(* IEC 61131-3 sources: iecf/harness/cases (part 2) *)

(* ---- enobody.st ---- *)
(* ENO set in a POU's own body (Ed.3 6.6.1.5 rules 2, 3 and 7;
   docs/dependencies.md): ENO is there in every FUNCTION and
   FUNCTION_BLOCK without a declaration, TRUE as each run starts, and the
   caller's ENO is FALSE when the body set it FALSE or a flag was raised
   while it ran. `lim` clears ENO above 100, `half` below 0; `acc` sets
   ENO TRUE at its end, which cannot hide the overflow of its fifth run
   (tick 4): iecf's ENO is FALSE there, the reference compiler's TRUE, as
   it has no flag; iecf's trace is enobody.iecf.trace. The input v is
   5, 200, -4, 30000, 30000. r_bits: bit 0 lim's ENO, 1 half's, 2 acc's. *)
FUNCTION_BLOCK lim
VAR_INPUT x : INT; END_VAR
VAR_OUTPUT y : INT; END_VAR
y := x;
IF x > 100 THEN ENO := FALSE; END_IF;
END_FUNCTION_BLOCK

FUNCTION half : INT
VAR_INPUT x : INT; END_VAR
half := x / 2;
ENO := x >= 0;
END_FUNCTION

FUNCTION_BLOCK acc
VAR_INPUT x : INT; END_VAR
VAR_OUTPUT total : INT; END_VAR
total := total + x;
ENO := TRUE;
END_FUNCTION_BLOCK

PROGRAM main
VAR
  v AT %IW0 : INT;
  r_bits AT %MB0 : BYTE;
  r_half AT %MB1 : SINT;
  r_y AT %MW2 : INT;
  r_total AT %MW4 : INT;
END_VAR
VAR
  l : lim;
  a : acc;
  ok1, ok2, ok3 : BOOL;
  h : INT;
END_VAR
l(x := v, y => r_y, ENO => ok1);
h := half(x := v, ENO => ok2);
r_half := INT_TO_SINT(h / 1000);
a(x := v, total => r_total, ENO => ok3);
r_bits := 0;
IF ok1 THEN r_bits := r_bits OR 16#01; END_IF;
IF ok2 THEN r_bits := r_bits OR 16#02; END_IF;
IF ok3 THEN r_bits := r_bits OR 16#04; END_IF;
END_PROGRAM

CONFIGURATION plant
  RESOURCE r ON PLC
    TASK fast(INTERVAL := T#10ms, PRIORITY := 0);
    PROGRAM p WITH fast : main;
  END_RESOURCE
END_CONFIGURATION

(* ---- enointo.st ---- *)
(* A block's ENO, and outputs, taken into an element, a field and a bit,
   each found - its index checked - before the block runs. Worked by
   hand:
   t(EN := TRUE, ..., ENO => a[i]), i 2: ENO TRUE, a[2] TRUE (%QX0.0).
   t(EN := FALSE, ..., NOT ENO => w.3): ENO FALSE, its NOT TRUE: w 8,
   w.%B0 08 (%QB1).
   t(EN := TRUE, ..., ENO => s.ok): s.ok TRUE (%QX0.1).
   o(q => ws[i].3, qb => ws[i].%B1), q TRUE and qb 7: ws[2] 16#0708,
   its bytes 08 (%QB2) and 07 (%QB3).
   F(q => ws[1].2), q TRUE: ws[1] 4 (%QB4).
   Last, i 3: o(q => ws[i].0) faults (INDEX) before o runs, so n, o's
   count of its runs, stays 1 (%QB5).
   reference-skip: partial access, NOT ENO =>: refused (iec2c crashes
   on the latter). *)
TYPE
  STV : STRUCT ok : BOOL; END_STRUCT;
END_TYPE
FUNCTION_BLOCK OT
  VAR_OUTPUT q : BOOL; qb : BYTE; n : INT; END_VAR
  q := TRUE;
  qb := 7;
  n := n + 1;
END_FUNCTION_BLOCK
FUNCTION F : INT
  VAR_OUTPUT q : BOOL; END_VAR
  q := TRUE;
  F := 1;
END_FUNCTION
PROGRAM main
  VAR
    t : TON;
    o : OT;
    a : ARRAY [1..2] OF BOOL;
    ws : ARRAY [1..2] OF WORD;
    s : STV;
    w : WORD;
    i : INT := 2;
    v : INT;
  END_VAR
  VAR
    q00 AT %QX0.0 : BOOL;
    q01 AT %QX0.1 : BOOL;
    q1 AT %QB1 : BYTE;
    q2 AT %QB2 : BYTE;
    q3 AT %QB3 : BYTE;
    q4 AT %QB4 : BYTE;
    q5 AT %QB5 : SINT;
  END_VAR
  t(EN := TRUE, IN := FALSE, PT := T#1s, ENO => a[i]);
  q00 := a[2];
  t(EN := FALSE, IN := FALSE, PT := T#1s, NOT ENO => w.3);
  q1 := w.%B0;
  t(EN := TRUE, IN := FALSE, PT := T#1s, ENO => s.ok);
  q01 := s.ok;
  o(q => ws[i].3, qb => ws[i].%B1);
  q2 := ws[2].%B0;
  q3 := ws[2].%B1;
  v := F(q => ws[1].2);
  q4 := ws[1].%B0;
  q5 := INT_TO_SINT(o.n);
  i := 3;
  o(q => ws[i].0);
END_PROGRAM

CONFIGURATION c
  RESOURCE r ON x
    TASK t(INTERVAL := T#10ms, PRIORITY := 1);
    PROGRAM p WITH t : main;
  END_RESOURCE
END_CONFIGURATION

(* ---- enums.st ---- *)
(* Enumerations and types with named values (Ed.3 6.4.4.2, 6.4.4.3).
   col has named values: red 1, green 5, blue one more, 6; its initial
   value green. A col is used as the INT it is: other values assigned,
   arithmetic, comparison. mode is an enumeration, its initial value run.
   An enumeration is a FUNCTION's input, output and result and a block's
   in-out; a result or an input not given starts as the type's initial
   value. Worked by hand, k %IB0 1, 2, 3:
   %QB0: c as the tick starts: 5 (green), then what the tick before left,
   3, 4. %QB1: x := c + blue when c = green: 11, and kept.
   c := k, then CASE c OF red: 10; green - 3 (2), blue: 20; ELSE 30:
   %QB2 10, 20, 30.
   b(c := c, m := m, d := red + 1): c + 2, %QB3 3, 4, 5; m := NEXT(m):
   run gives stop; stop matches no label, so NEXT keeps its initial value,
   run; then stop again: %QB4 2, 1, 2 (stop 2, run 1).
   lv#hi OR lo, a WORD: 16#30, %QB5.
   n, an INT, given to the in-out c: 10 + blue each tick: %QB6 16, 22, 28.
   m3 := DEF(o => m4), both idle before: DEF's result is not set and its
   input m not given, so both are run: %QB7 1.
   %QB8 blue, 6. %QB9 a[2], an array's element of col: green, 5.
   mi : (low, mid, top) := mid, declared in place: mid gives 7 and
   becomes top, top gives 8: %QB10 7, 8, 8.
   gear names no base type, so it is an INT (as CODESYS and TwinCAT
   have it) and is added to one as it is: g is slow, 2; x2, an INT from
   3, x2 := x2 + g each tick: %QB11 5, 7, 9.
   reference-skip: named values are Ed.3's; the reference compiler
   (Ed.2) has none. *)
TYPE
  col : INT (red := 1, green := 5, blue) := green;
  lv : WORD (lo := 16#10, hi := 16#20);
  mode : (idle, run, stop) := run;
  gear : (slow := 2, fast := 4);
END_TYPE

FUNCTION NEXT : mode
  VAR_INPUT m : mode; END_VAR
  CASE m OF
    idle: NEXT := run;
    run: NEXT := stop;
  END_CASE;
END_FUNCTION

FUNCTION DEF : mode
  VAR_INPUT m : mode; END_VAR
  VAR_OUTPUT o : mode; END_VAR
  o := m;
END_FUNCTION

FUNCTION_BLOCK BUMP
  VAR_IN_OUT c : col; m : mode; END_VAR
  VAR_INPUT d : col; END_VAR
  c := c + d;
  m := NEXT(m);
END_FUNCTION_BLOCK

PROGRAM main
  VAR
    c : col;
    x : INT;
    w : WORD;
    m, m2 : mode;
    m3, m4 : mode := idle;
    b : BUMP;
    n : INT := 10;
    a : ARRAY [1..2] OF col;
    mi : (low, mid, top) := mid;
    g : gear;
    x2 : INT := 3;
  END_VAR
  VAR k AT %IB0 : SINT; END_VAR
  VAR
    q0 AT %QB0 : SINT;
    q1 AT %QB1 : SINT;
    q2 AT %QB2 : SINT;
    q3 AT %QB3 : SINT;
    q4 AT %QB4 : SINT;
    q5 AT %QB5 : BYTE;
    q6 AT %QB6 : SINT;
    q7 AT %QB7 : SINT;
    q8 AT %QB8 : SINT;
    q9 AT %QB9 : SINT;
    q10 AT %QB10 : SINT;
    q11 AT %QB11 : SINT;
  END_VAR
  q0 := INT_TO_SINT(c);
  IF c = col#green THEN
    x := c + blue;
  END_IF;
  q1 := INT_TO_SINT(x);
  c := k;
  CASE c OF
    red: q2 := 10;
    green - 3, blue: q2 := 20;
  ELSE
    q2 := 30;
  END_CASE;
  b(c := c, m := m, d := red + 1);
  q3 := INT_TO_SINT(c);
  IF m = stop THEN
    q4 := 2;
  ELSIF m = mode#run THEN
    q4 := 1;
  ELSE
    q4 := 0;
  END_IF;
  w := lv#hi OR lo;
  q5 := WORD_TO_BYTE(w);
  b(c := n, m := m2, d := blue);
  q6 := INT_TO_SINT(n);
  m3 := DEF(o => m4);
  IF m3 = run AND m4 = run THEN
    q7 := 1;
  END_IF;
  q8 := INT_TO_SINT(blue);
  q9 := INT_TO_SINT(a[2]);
  IF mi = mid THEN
    q10 := 7;
    mi := top;
  ELSIF mi = top THEN
    q10 := 8;
  END_IF;
  x2 := x2 + g;
  q11 := INT_TO_SINT(x2);
END_PROGRAM

CONFIGURATION c
  RESOURCE r ON PLC
    TASK t(INTERVAL := T#10ms, PRIORITY := 1);
    PROGRAM p WITH t : main;
  END_RESOURCE
END_CONFIGURATION

(* ---- fbargs.st ---- *)
(* A function block's in-out given, and its output taken into, any
   variable of the type (Ed.3 6.6.3.4): an element by a constant and by
   a computed index, a field, a variable through a reference, an
   element at an address. And an enumeration declared in place with
   named values (Ed.3 6.4.4.3), used as its base type.
   ADD1 adds 1 to its in-out v; twice := 2 * v; neg := v < 0.
   Worked by hand, k %IB0 1, 2, 3; arr and out start [0, 0, 0]:
   b(v := arr[2], twice => out[1]); i := k; b(v := arr[i], twice =>
   out[i]); and, last in the scan, b(v := arr[k + 1]):
     tick 0: arr[2] 1, out[1] 2; i 1: arr[1] 1, out[1] 2; arr [1, 1,
     0], out [2, 0, 0]; then arr[2] 2.
     tick 1: arr[2] 3, out[1] 6; i 2: arr[2] 4, out[2] 8; arr [1, 4,
     0], out [6, 8, 0]; then arr[3] 1.
     tick 2: arr[2] 5, out[1] 10; i 3: arr[3] 2, out[3] 4; arr [1, 5,
     2], out [10, 8, 4]; then arr[4], outside 1..3: a fault (index),
     before the block runs.
     %QB0..2 arr, %QB3..5 out.
   b(v := p.y, twice => po.x): p.y 1, 2, 3 (%QB6); po.x 2, 4, 6 (%QB7).
   b(v := r^, twice => ro^), r to tgt, ro to d2: tgt + 1, d2 twice it.
   b(v := tgt, twice => d), d a DINT, the output widened: tgt + 1
   again: tgt 2, 4, 6 (%QB8); d2 2, 6, 10 (%QB9); d 4, 8, 12 (%QB10).
   b(v := p.x, NOT neg => nb): nb TRUE (%QX11.0).
   b(v := lm[2], twice => lm[1]), lm at %MW0: lm[2] 1, 2, 3 and lm[1]
   2, 4, 6 in %MW2 and %MW0.
   x : INT (lo := 1, hi := 5) := hi, in place: x + lo 6, then x := x + 1:
   6, 7, 8 (%QB12). y : (p3 := 3, q4): 3, then y := q4: 3, 4, 4 (%QB13).
   SPARE is a block with an instance that is never called: the C still
   builds with every warning an error, as the harness builds it.
   reference-skip: named values are Ed.3's; the reference compiler
   (Ed.2) has none. *)
TYPE PT : STRUCT x, y : INT; END_STRUCT; END_TYPE
FUNCTION_BLOCK ADD1
  VAR_IN_OUT v : INT; END_VAR
  VAR_OUTPUT twice : INT; neg : BOOL; END_VAR
  v := v + 1;
  twice := 2 * v;
  neg := v < 0;
END_FUNCTION_BLOCK
FUNCTION_BLOCK SPARE
  VAR_INPUT a : INT; END_VAR
  VAR_OUTPUT o : INT; END_VAR
  o := a;
END_FUNCTION_BLOCK
CONFIGURATION c
  RESOURCE r ON PLC
    TASK t(INTERVAL := T#10ms, PRIORITY := 1);
    PROGRAM p WITH t : main;
  END_RESOURCE
END_CONFIGURATION
PROGRAM main
  VAR
    arr, out : ARRAY [1..3] OF INT;
    p, po : PT;
    r, ro : REF_TO INT;
    tgt, d2, i : INT;
    d : DINT;
    nb : BOOL;
    b : ADD1;
    idle : SPARE;
    x : INT (lo := 1, hi := 5) := hi;
    y : (p3 := 3, q4);
  END_VAR
  VAR lm AT %MW0 : ARRAY [1..2] OF INT; END_VAR
  VAR k AT %IB0 : SINT; END_VAR
  VAR
    q0 AT %QB0 : SINT;
    q1 AT %QB1 : SINT;
    q2 AT %QB2 : SINT;
    q3 AT %QB3 : SINT;
    q4b AT %QB4 : SINT;
    q5 AT %QB5 : SINT;
    q6 AT %QB6 : SINT;
    q7 AT %QB7 : SINT;
    q8 AT %QB8 : SINT;
    q9 AT %QB9 : SINT;
    q10 AT %QB10 : SINT;
    q11 AT %QX11.0 : BOOL;
    q12 AT %QB12 : SINT;
    q13 AT %QB13 : SINT;
  END_VAR
  b(v := arr[2], twice => out[1]);
  i := k;
  b(v := arr[i], twice => out[i]);
  b(v := p.y, twice => po.x);
  r := REF(tgt);
  ro := REF(d2);
  b(v := r^, twice => ro^);
  b(v := tgt, twice => d);
  b(v := p.x, NOT neg => nb);
  b(v := lm[2], twice => lm[1]);
  q0 := INT_TO_SINT(arr[1]);
  q1 := INT_TO_SINT(arr[2]);
  q2 := INT_TO_SINT(arr[3]);
  q3 := INT_TO_SINT(out[1]);
  q4b := INT_TO_SINT(out[2]);
  q5 := INT_TO_SINT(out[3]);
  q6 := INT_TO_SINT(p.y);
  q7 := INT_TO_SINT(po.x);
  q8 := INT_TO_SINT(tgt);
  q9 := INT_TO_SINT(d2);
  q10 := DINT_TO_SINT(d);
  q11 := nb;
  q12 := INT_TO_SINT(x + lo);
  x := x + 1;
  q13 := INT_TO_SINT(y);
  y := q4;
  b(v := arr[k + 1]);
END_PROGRAM

(* ---- fbeffects.st ---- *)
(* FUNCTIONs with effects in a block call: in the index of the target an
   output is taken into, and as a STRING input. Each is made once, in
   order; an output's target is found after the block runs, as a
   FUNCTION's is, so a call there runs after the block does
   (docs/dependencies.md). Worked by hand, each tick from j 1:

   f(io := j, s := 'x', q => a[finc(j)]): the block, io j 1: q 1 +
   LEN('x') 1 = 2; then finc makes j 2 and gives 2, the target a[2]:
   2 (Q0 02). f(io := j, s := fso(x := 'bb', y => j)): fso gives
   'bb' and sets j to 7; then the block, io 7: q 7 + 2 = 9 (Q1 09); j 7
   (Q2 07).
   fbeffects.iecf.trace: the reference compiler copies the in-out in
   before the other inputs are computed and back after the call, so
   fso's j is lost (Q 02 04 02); iecf binds the in-out to j itself. *)
FUNCTION finc : INT
  VAR_IN_OUT x : INT; END_VAR
  x := x + 1;
  finc := x;
END_FUNCTION
FUNCTION fso : STRING
  VAR_INPUT x : STRING; END_VAR
  VAR_OUTPUT y : INT; END_VAR
  y := 7;
  fso := x;
END_FUNCTION
FUNCTION_BLOCK fb
  VAR_IN_OUT io : INT; END_VAR
  VAR_INPUT s : STRING; END_VAR
  VAR_OUTPUT q : INT; END_VAR
  q := io + LEN(s);
END_FUNCTION_BLOCK
PROGRAM main
  VAR f : fb; a : ARRAY [1..4] OF INT; j : INT; END_VAR
  VAR q AT %QB0 : USINT; q1 AT %QB1 : USINT; q2 AT %QB2 : USINT; END_VAR
  j := 1;
  f(io := j, s := 'x', q => a[finc(j)]);
  q := INT_TO_USINT(a[2]);
  f(io := j, s := fso(x := 'bb', y => j));
  q1 := INT_TO_USINT(f.q);
  q2 := INT_TO_USINT(j);
END_PROGRAM
CONFIGURATION c RESOURCE r ON PLC TASK t(INTERVAL := T#10ms, PRIORITY := 1); PROGRAM p WITH t : main; END_RESOURCE END_CONFIGURATION

(* ---- fbenable.st ---- *)
(* EN and ENO on a function block call (Ed.3 6.6.1.5; docs/dependencies.md):
   an accumulator adds 10000 at each call it is enabled for, %IX0.0 its EN.
   Each tick r_n is set to -1 before the call: with EN FALSE (tick 1) the
   block is not called, its total stays and is not taken into r_n, and ENO
   is FALSE. Its fourth enabled call (tick 4) overflows inside the block:
   the total wraps, the flag is raised in the block's body, and ENO is
   FALSE. r_bits: bit 0 ENO. The reference compiler takes the output into
   r_n with EN FALSE and has no flag to clear ENO: iecf's trace is
   fbenable.iecf.trace. NOT ENO, which the reference compiler cannot
   compile, is fbskip's. *)
FUNCTION_BLOCK acc
VAR_INPUT x : INT; END_VAR
VAR_OUTPUT total : INT; END_VAR
total := total + x;
END_FUNCTION_BLOCK

PROGRAM main
VAR
  c AT %IX0.0 : BOOL;
  r_n AT %MW0 : INT;
  r_total AT %MW2 : INT;
  r_bits AT %MB4 : BYTE;
END_VAR
VAR
  a : acc;
  ok : BOOL;
END_VAR
r_n := -1;
a(EN := c, x := 10000, total => r_n, ENO => ok);
r_total := a.total;
r_bits := 0;
IF ok THEN r_bits := r_bits OR 16#01; END_IF;
END_PROGRAM

CONFIGURATION plant
  RESOURCE r ON PLC
    TASK fast(INTERVAL := T#10ms, PRIORITY := 0);
    PROGRAM p WITH fast : main;
  END_RESOURCE
END_CONFIGURATION

(* ---- fbencall.st ---- *)
(* A function block's EN given a call (Ed.3 6.6.1.5): of a FUNCTION
   with an in-out, of a method, of a method through an interface. EN is
   computed first, once, and only then the block is called or not, ENO
   telling which. Worked by hand, tick by tick:
   Advance adds 1 to n and gives n > 2: n 1, 2, 3, 4; c1 runs at ticks
   2 and 3, total (%QB0) 0, 0, 1, 2; n (%QB1); ENO e1 (%QX4.0) FALSE,
   FALSE, TRUE, TRUE.
   v.Ready gives its count < 2, then counts: TRUE, TRUE, FALSE, FALSE;
   c2 adds 10: 10, 20, 20, 20 (%QB2); e2 (%QX4.1).
   ig.Open counts and gives whether its count is even: FALSE, TRUE,
   FALSE, TRUE; c3 adds 5: 0, 5, 5, 10 (%QB3); e3 (%QX4.2).
   reference-skip: METHOD and INTERFACE are Ed.3's; the reference
   compiler (Ed.2) has neither. *)
FUNCTION Advance : BOOL
  VAR_IN_OUT cnt : INT; END_VAR
  cnt := cnt + 1;
  Advance := cnt > 2;
END_FUNCTION

FUNCTION_BLOCK Valve
  VAR n : INT; END_VAR
  METHOD PUBLIC Ready : BOOL
    Ready := n < 2;
    n := n + 1;
  END_METHOD
END_FUNCTION_BLOCK

INTERFACE IGate
  METHOD Open : BOOL
  END_METHOD
END_INTERFACE

FUNCTION_BLOCK Gate IMPLEMENTS IGate
  VAR k : INT; END_VAR
  METHOD PUBLIC Open : BOOL
    k := k + 1;
    Open := k MOD 2 = 0;
  END_METHOD
END_FUNCTION_BLOCK

FUNCTION_BLOCK Count
  VAR_INPUT inc : INT; END_VAR
  VAR_OUTPUT total : INT; END_VAR
  total := total + inc;
END_FUNCTION_BLOCK

PROGRAM main
  VAR
    n : INT;
    v : Valve;
    g : Gate;
    ig : IGate;
    c1, c2, c3 : Count;
  END_VAR
  VAR
    q0 AT %QB0 : SINT;
    q1 AT %QB1 : SINT;
    q2 AT %QB2 : SINT;
    q3 AT %QB3 : SINT;
    e1 AT %QX4.0 : BOOL;
    e2 AT %QX4.1 : BOOL;
    e3 AT %QX4.2 : BOOL;
  END_VAR
  ig := g;
  c1(EN := Advance(n), inc := 1, ENO => e1);
  c2(EN := v.Ready(), inc := 10, ENO => e2);
  c3(EN := ig.Open(), inc := 5, ENO => e3);
  q0 := INT_TO_SINT(c1.total);
  q1 := INT_TO_SINT(n);
  q2 := INT_TO_SINT(c2.total);
  q3 := INT_TO_SINT(c3.total);
END_PROGRAM

CONFIGURATION c
  RESOURCE r ON x
    TASK t(INTERVAL := T#10ms, PRIORITY := 1);
    PROGRAM p WITH t : main;
  END_RESOURCE
END_CONFIGURATION

(* ---- fbinitarrays.st ---- *)
(* CODESYS's and TwinCAT's arrays of instances set up by their FB_init
   (fb-init), as TcOpen's `ARRAY[0..2] OF DiagnosticsMessenger(THIS^)`,
   and in-outs of a type with an FB_init, bound, not set up.
   Worked by hand: h's items, its first VAR, are set up first, each
   element's FB_init in index order given THIS^, h: each takes h.Next(),
   1 2 3; then grid, row by row, (1,-1) (1,0) (2,-1) (2,0): 4 5 6 7;
   then plain, with no arguments, each element's FB_init counting itself
   once, bInitRetains TRUE at the cold start; then d, a structure whose
   member cells is such an array, then nest, an array of arrays.
   %QW0 items[0..2] 1 2 3 as 123, %QW2 grid as 4567, %QW4 h.seq 7,
   %QW6 plain's counts summed, 3, %QW8 those cold, 3, %QW10 d.cells'
   counts summed, 2, and nest's, 4, times 10: 42; %QW12 h.u reading items[2] through its in-out, 3,
   %QW14 its method reading grid[2, 0] through one, 7.
   reference-skip: not IEC 61131-3. *)
INTERFACE ISeq
  METHOD Next : INT
  END_METHOD
END_INTERFACE

FUNCTION_BLOCK Item
  VAR_OUTPUT mine : INT; END_VAR
  METHOD FB_init : BOOL
    VAR_INPUT bInitRetains : BOOL; bInCopyCode : BOOL; s : ISeq; END_VAR
    mine := s.Next();
  END_METHOD
END_FUNCTION_BLOCK

FUNCTION_BLOCK Counted
  VAR_OUTPUT times : INT; cold : INT; END_VAR
  METHOD FB_init : BOOL
    VAR_INPUT bInitRetains : BOOL; bInCopyCode : BOOL; END_VAR
    times := times + 1;
    IF bInitRetains THEN cold := cold + 1; END_IF
  END_METHOD
END_FUNCTION_BLOCK

TYPE Cells : STRUCT
  tag : INT := 1;
  cells : ARRAY[0..1] OF Counted;
END_STRUCT
END_TYPE

FUNCTION_BLOCK User
  VAR_IN_OUT io : Item; END_VAR
  VAR_OUTPUT o : INT; END_VAR
  METHOD Read : INT
    VAR_IN_OUT other : Item; END_VAR
    Read := other.mine;
  END_METHOD
  o := io.mine;
END_FUNCTION_BLOCK

FUNCTION_BLOCK Holder IMPLEMENTS ISeq
  VAR
    seq : INT;
    items : ARRAY[0..2] OF Item(THIS^);
    grid : ARRAY[1..2, -1..0] OF Item(THIS^);
    plain : ARRAY[0..2] OF Counted;
    d : Cells;
    nest : ARRAY[0..1] OF ARRAY[0..1] OF Counted;
    u : User;
  END_VAR
  VAR_OUTPUT o1 : INT; o2 : INT; o3 : INT; o4 : INT; o5 : INT; o6 : INT; o7 : INT; o8 : INT; END_VAR
  VAR_TEMP k : INT; END_VAR
  METHOD PUBLIC Next : INT
    seq := seq + 1;
    Next := seq;
  END_METHOD
  o1 := items[0].mine * 100 + items[1].mine * 10 + items[2].mine;
  o2 := grid[1, -1].mine * 1000 + grid[1, 0].mine * 100 + grid[2, -1].mine * 10 + grid[2, 0].mine;
  o3 := seq;
  o4 := 0; o5 := 0;
  FOR k := 0 TO 2 DO
    o4 := o4 + plain[k].times;
    o5 := o5 + plain[k].cold;
  END_FOR
  o6 := d.cells[0].times + d.cells[1].times;
  FOR k := 0 TO 1 DO
    o6 := o6 + 10 * (nest[k][0].times + nest[k][1].times);
  END_FOR
  u(io := items[2]);
  o7 := u.o;
  o8 := u.Read(other := grid[2, 0]);
END_FUNCTION_BLOCK

PROGRAM main
  VAR h : Holder; END_VAR
  VAR q0 AT %QW0 : INT; q1 AT %QW2 : INT; q2 AT %QW4 : INT; q3 AT %QW6 : INT; q4 AT %QW8 : INT;
      q5 AT %QW10 : INT; q6 AT %QW12 : INT; q7 AT %QW14 : INT; END_VAR
  h();
  q0 := h.o1; q1 := h.o2; q2 := h.o3; q3 := h.o4; q4 := h.o5; q5 := h.o6;
  q6 := h.o7; q7 := h.o8;
END_PROGRAM

CONFIGURATION cf
  RESOURCE r ON x
    TASK tk(INTERVAL := T#10ms, PRIORITY := 1);
    PROGRAM p WITH tk : main;
  END_RESOURCE
END_CONFIGURATION

(* ---- fbinorder.st ---- *)
(* A function block called with its arguments in order (Ed.3 6.6.3.4.1,
   the non-formal call): every input, output and in-out where it is
   declared, a base's first, none left off ("exactly the same number of
   parameters, in exactly the same order", 6.6.1.4.2). Worked by hand:

   tick 0. adder declares a, b, o, n, o2: f(1, 2, r, x, r2) gives a 1,
   b 2, o into r, the in-out n is x, o2 into r2: r 3 (Q0), r2 -1 (Q2 ff
   ff), x 1 (Q4). f(10, 20, r, x, r2): f.o 30 (Q6 1e 00), x 2. g, a
   wider, takes adder's a, b, o, n, o2, then its own c, p, s, o3: g(1,
   2, r, x, r2, 3, pt, 'abc', r3) gives o 3, x 3, o3 3 + 3 + 100 + 3 =
   109 (Q8 6d 00). g.twice(7, h): 14, h 3: 17 (Q10 11 00). TON's IN,
   PT, Q, ET: t(TRUE, T#20ms, done, el): not done (Q12 0); CTU's CU, R,
   PV, Q, CV: ctr(done, FALSE, 5, cq, cv): 0 (Q14).
   tick 1: x was 3: 4 after the first call (Q4 04 00); the rest as
   before.
   tick 2: x 7; t is done after 20 ms (Q12 01 00), and ctr counts its
   rising edge: 1 (Q14).
   tick 3: x 10; done stays, the count stays 1.
   reference-skip: methods, EXTENDS: refused. *)
TYPE PtT : STRUCT x : INT; y : INT; END_STRUCT; END_TYPE
FUNCTION_BLOCK adder
  VAR_INPUT a : INT; b : INT := 5; END_VAR
  VAR_OUTPUT o : INT; END_VAR
  VAR_IN_OUT n : INT; END_VAR
  VAR_OUTPUT o2 : INT; END_VAR
  o := a + b;
  n := n + 1;
  o2 := a - b;
END_FUNCTION_BLOCK
FUNCTION_BLOCK wider EXTENDS adder
  VAR_INPUT c : INT; p : PtT; s : STRING[4]; END_VAR
  VAR_OUTPUT o3 : INT; END_VAR
  METHOD PUBLIC twice : INT
    VAR_INPUT v : INT; END_VAR
    VAR_OUTPUT half : INT; END_VAR
    twice := v * 2;
    half := v / 2;
  END_METHOD
  SUPER();
  o3 := o + c + p.x + LEN(s);
END_FUNCTION_BLOCK
PROGRAM main
  VAR f : adder; g : wider; t : TON; ctr : CTU; x : INT; r, r2, r3, m, h : INT; pt : PtT := (x := 100); el : TIME; done, cq : BOOL; cv : INT; END_VAR
  VAR q AT %QW0 : ARRAY [0..7] OF INT; END_VAR
  f(1, 2, r, x, r2);
  q[0] := r; q[1] := r2; q[2] := x;
  f(10, 20, r, x, r2);
  q[3] := f.o;
  g(1, 2, r, x, r2, 3, pt, 'abc', r3);
  q[4] := r3;
  m := g.twice(7, h);
  q[5] := m + h;
  t(TRUE, T#20ms, done, el);
  q[6] := BOOL_TO_INT(done);
  ctr(done, FALSE, 5, cq, cv);
  q[7] := ctr.CV;
END_PROGRAM
CONFIGURATION c RESOURCE r ON PLC TASK t(INTERVAL := T#10ms, PRIORITY := 1); PROGRAM p WITH t : main; END_RESOURCE END_CONFIGURATION

(* ---- fbparts.st ---- *)
(* A part of a block's elementary input or output read from outside
   (Ed.3 Table 17): `f.q.%X4`, `f.q.%B1`, of an element of an array of
   instances, in a condition. Worked by hand: f.iw 16#0123, so f.q is
   ROL(16#0123, 4), 16#1230: its byte 1 is 16#12 (Q0); its bit 4 is 1,
   iw's bit 1 is 1, fa[2].q is 16#0040 and its bit 6 is 1, f.q's bit 5
   is 1: the four bits 2#1111 (Q1 0f).
   reference-skip: partial access, as `partaccess`. *)
FUNCTION_BLOCK fb
  VAR_INPUT iw : WORD; END_VAR
  VAR_OUTPUT q : WORD; END_VAR
  q := ROL(iw, 4);
END_FUNCTION_BLOCK
PROGRAM main
  VAR f : fb; fa : ARRAY [1..2] OF fb; i : INT := 2; b1, b2, b3, b4 : BOOL; y : BYTE; END_VAR
  VAR q AT %QB0 : BYTE; q1 AT %QB1 : BYTE; END_VAR
  f(iw := 16#0123);
  fa[2](iw := 16#0004);
  b1 := f.q.%X4;
  y := f.q.%B1;
  b2 := f.iw.%X1;
  b3 := fa[i].q.%X6;
  IF f.q.%X5 THEN b4 := TRUE; END_IF;
  q := y;
  q1 := BOOL_TO_BYTE(b1) OR SHL(BOOL_TO_BYTE(b2), 1) OR SHL(BOOL_TO_BYTE(b3), 2) OR SHL(BOOL_TO_BYTE(b4), 3);
END_PROGRAM
CONFIGURATION c RESOURCE r ON PLC TASK t(INTERVAL := T#10ms, PRIORITY := 1); PROGRAM p WITH t : main; END_RESOURCE END_CONFIGURATION

(* ---- fbretain.st ---- *)
(* RETAIN inside a FUNCTION_BLOCK (Ed.3 6.5.6): at a warm restart the
   block's own RETAIN variable keeps its value, its NON_RETAIN one is set
   anew, and one that is neither keeps its value only in an instance
   declared RETAIN. A block in a block follows its own type and the
   section it is declared in, not the outer instance. An instance of a
   block that keeps anything is kept whole (docs/c-output.md §7).
   Each counter counts from 10, 20, 30; at tick 3 a warm restart.
   The reference compiler has no warm restart of its own; its host starts everything
   anew. iecf's trace is fbretain.iecf.trace. *)
FUNCTION_BLOCK cnt
VAR_OUTPUT
  ko : INT;
  po : INT;
  no : INT;
END_VAR
VAR RETAIN
  k : INT := 10;
END_VAR
VAR
  p : INT := 20;
END_VAR
VAR NON_RETAIN
  n : INT := 30;
END_VAR
k := k + 1;
p := p + 1;
n := n + 1;
ko := k;
po := p;
no := n;
END_FUNCTION_BLOCK

FUNCTION_BLOCK wrap
VAR_OUTPUT
  ck, cp, cn, dk, dp, dn : INT;
END_VAR
VAR
  c : cnt;
END_VAR
VAR RETAIN
  cr : cnt;
END_VAR
c();
cr();
ck := c.ko;
cp := c.po;
cn := c.no;
dk := cr.ko;
dp := cr.po;
dn := cr.no;
END_FUNCTION_BLOCK

PROGRAM main
VAR
  a_k AT %MW0 : INT;
  a_p AT %MW2 : INT;
  a_n AT %MW4 : INT;
  b_k AT %MW6 : INT;
  b_p AT %MW8 : INT;
  b_n AT %MW10 : INT;
  c_k AT %MW12 : INT;
  c_p AT %MW14 : INT;
  c_n AT %MW16 : INT;
  d_k AT %MW18 : INT;
  d_p AT %MW20 : INT;
  d_n AT %MW22 : INT;
END_VAR
VAR
  a : cnt;
  w : wrap;
END_VAR
VAR RETAIN
  b : cnt;
END_VAR
a();
b();
w();
a_k := a.ko;
a_p := a.po;
a_n := a.no;
b_k := b.ko;
b_p := b.po;
b_n := b.no;
c_k := w.ck;
c_p := w.cp;
c_n := w.cn;
d_k := w.dk;
d_p := w.dp;
d_n := w.dn;
END_PROGRAM

CONFIGURATION plant
  RESOURCE r ON PLC
    TASK fast(INTERVAL := T#10ms, PRIORITY := 0);
    PROGRAM p WITH fast : main;
  END_RESOURCE
END_CONFIGURATION

(* ---- fbskip.st ---- *)
(* A function block call with EN FALSE is not made at all (Ed.3 6.6.1.5,
   Example 2; docs/dependencies.md): its inputs are not evaluated - x
   divides by zero and nothing faults - nor set, the block does not run,
   its output is not taken, and NOT ENO gives TRUE. With EN TRUE at tick 1
   (zero is 1 by then) it runs once. The reference compiler cannot compile
   `NOT ENO =>` (PROPOSAL.md §1b): iecf only. *)
FUNCTION_BLOCK acc
VAR_INPUT x : INT; END_VAR
VAR_OUTPUT total : INT; END_VAR
total := total + x;
END_FUNCTION_BLOCK

PROGRAM main
VAR
  r_n AT %MW0 : INT;
  r_total AT %MW2 : INT;
  r_off AT %MX4.0 : BOOL;
END_VAR
VAR
  a : acc;
  run : BOOL;
  zero : INT;
END_VAR
r_n := -1;
a(EN := run, x := 100 / zero, total => r_n, NOT ENO => r_off);
r_total := a.total;
run := TRUE;
zero := 1;
END_PROGRAM

CONFIGURATION plant
  RESOURCE r ON PLC
    TASK fast(INTERVAL := T#10ms, PRIORITY := 0);
    PROGRAM p WITH fast : main;
  END_RESOURCE
END_CONFIGURATION

(* ---- flexarrays.st ---- *)
(* Variable-length arrays (Ed.3 6.5.3) and named constants in bounds
   (Ed.3 6.6.1.2.4). SUM is Ed.3's Example 2: it adds an ARRAY[*] whatever
   its bounds. FILL writes a 2-dimensional one, M[i, j] := 10 * i + j.
   TWICE passes its ARRAY[*] on to SUM. A CLASS's method takes one too.
   W, a VAR_GLOBAL CONSTANT, bounds a TYPE; N, the program's own
   CONSTANT, bounds an array and a STRING; a subrange is 0..N.
   Worked by hand, k %IB0:
   a: 1..5 (N), [1, 2, 3, 4, 5]: SUM 15, %QB0 15. b: -2..2, [10, 20, 30,
   40, 50]: SUM 150, %QB1 150. TWICE(a) 2 * 15 = 30, %QB2 30.
   m: 1..2, -1..1 filled: m[1, -1] 9, m[2, 1] 21: %QB3 9, %QB4 21.
   LOWER_BOUND(b, 1) -2, %QB5 16#fe; UPPER_BOUND(m, 2) 1, %QB6 1.
   row: RowT, 0..W (W 3), [1, 1, 1, 1]: the method's COUNT gives 4,
   %QB7 4. LEN(s), s : STRING[N] := 'abcde': %QB8 5.
   lim : INT(0..N) := N: %QB9 5.
   Each tick, %QB10 := UPPER_BOUND(m, k): k 1 at tick 0, 2; k 2 at
   tick 1, 1. At tick 2, k 3: m has 2 dimensions, a fault (index), the
   statement stopped and %QB10 kept 1.
   A FUNCTION_BLOCK's in-outs, set by each call before the statement
   that faults: sc doubles c's elements, an ARRAY[*] ([1, 2, 3] at 0..2):
   c[2] 6, 12, 24 at ticks 0, 1, 2 (%QB11); f[2] := f[1] + f[3], 5
   (%QB12); t := CONCAT(t, 'x') on st, 'ab': LEN 3, 4, 5 (%QB13); p.a
   + 1 on pr: 1, 2, 3 (%QB14).
   A CASE's labels are constant expressions too (Ed.3 7.3.3.3.3): N - 4
   is 1, 2..W - 1 is 2..2: k 1, 2, 3 give %QB15 10, 20 and the ELSE's 30.
   A row of an array of arrays is an array (Ed.3 Example 2's SUM(A2[2])
   on the form the vendors take, docs/dependencies.md): aa, [[1, 2, 3],
   [4, 5, 6]]: SUM(aa[2]) 15 (%QB16); SUM(aa[k MOD 2 + 1]), the row
   computed: rows 2, 1, 2, so 15, 6, 15 (%QB17).
   An array of two dimensions indexed in the first only is the array of
   the second, Example 2's SUM(A2[2]) as written. m filled is [[9, 10,
   11], [19, 20, 21]]: SUM(m[2]) 60 (%QB18); SUM(m[k MOD 2 + 1]), rows
   2, 1, 2: 60, 30, 60 (%QB19). r3 := m[1] copies a row: r3[1] 11
   (%QB20). ROWSUM takes an ARRAY[*, *] and gives SUM(M[i]), a part of
   an ARRAY[*] passed on: ROWSUM(m, 1) 30 (%QB21).
   A row of an array at an address: lm at %MW0, 2 by 3 INTs; lm[2] :=
   r3 writes 9, 10, 11 at %MW6, %MW8, %MW10, the first row left 0; r4
   := lm[2] reads it back: r4[0] 10 (%QB22).
   reference-skip: ARRAY[*], LOWER_BOUND and UPPER_BOUND are Ed.3's, and
   CLASS; the reference compiler (Ed.2) has none. *)
TYPE RowT : ARRAY [0..W] OF SINT; END_TYPE
TYPE PAIR : STRUCT a : SINT; b : SINT; END_STRUCT; END_TYPE

FUNCTION_BLOCK SCALE
  VAR_INPUT k : INT; END_VAR
  VAR_IN_OUT
    v : ARRAY [*] OF INT;
    f : ARRAY [1..3] OF INT;
    t : STRING[5];
    p : PAIR;
  END_VAR
  VAR i : DINT; END_VAR
  FOR i := LOWER_BOUND(v, 1) TO UPPER_BOUND(v, 1) DO
    v[i] := v[i] * k;
  END_FOR;
  f[2] := f[1] + f[3];
  t := CONCAT(t, 'x');
  p.a := p.a + 1;
END_FUNCTION_BLOCK

FUNCTION SUM : DINT
  VAR_IN_OUT A : ARRAY [*] OF INT; END_VAR
  VAR i, s : DINT; END_VAR
  s := 0;
  FOR i := LOWER_BOUND(A, 1) TO UPPER_BOUND(A, 1) DO
    s := s + A[i];
  END_FOR;
  SUM := s;
END_FUNCTION

FUNCTION TWICE : DINT
  VAR_IN_OUT A : ARRAY [*] OF INT; END_VAR
  TWICE := 2 * SUM(A);
END_FUNCTION

FUNCTION ROWSUM : DINT
  VAR_IN_OUT M : ARRAY [*, *] OF INT; END_VAR
  VAR_INPUT i : INT; END_VAR
  ROWSUM := SUM(M[i]);
END_FUNCTION
FUNCTION FILL
  VAR_IN_OUT M : ARRAY [*, *] OF INT; END_VAR
  VAR i, j : DINT; END_VAR
  FOR i := LOWER_BOUND(ARR := M, DIM := 1) TO UPPER_BOUND(ARR := M, DIM := 1) DO
    FOR j := LOWER_BOUND(M, 2) TO UPPER_BOUND(M, 2) DO
      M[i, j] := DINT_TO_INT(10 * i + j);
    END_FOR;
  END_FOR;
END_FUNCTION

CLASS COUNTER
  METHOD PUBLIC COUNT : SINT
    VAR_IN_OUT r : ARRAY [*] OF SINT; END_VAR
    VAR i : DINT; END_VAR
    COUNT := 0;
    FOR i := LOWER_BOUND(r, 1) TO UPPER_BOUND(r, 1) DO
      COUNT := COUNT + r[i];
    END_FOR;
  END_METHOD
END_CLASS

CONFIGURATION c
  VAR_GLOBAL CONSTANT W : INT := 3; END_VAR
  RESOURCE r ON PLC
    TASK t(INTERVAL := T#10ms, PRIORITY := 1);
    PROGRAM p WITH t : main;
  END_RESOURCE
END_CONFIGURATION

PROGRAM main
  VAR CONSTANT N : INT := 5; END_VAR
  VAR_EXTERNAL CONSTANT W : INT; END_VAR
  VAR
    a : ARRAY [1..N] OF INT := [1, 2, 3, 4, 5];
    b : ARRAY [-2..2] OF INT := [10, 20, 30, 40, 50];
    m : ARRAY [1..2, -1..1] OF INT;
    row : RowT := [4(1)];
    cnt : COUNTER;
    s : STRING[N] := 'abcde';
    lim : INT (0..N) := N;
    c : ARRAY [0..2] OF INT := [1, 2, 3];
    f : ARRAY [1..3] OF INT := [1, 0, 4];
    st : STRING[5] := 'ab';
    pr : PAIR;
    sc : SCALE;
    aa : ARRAY [1..2] OF ARRAY [0..2] OF INT := [[1, 2, 3], [4, 5, 6]];
    r3 : ARRAY [-1..1] OF INT;
    r4 : ARRAY [-1..1] OF INT;
  END_VAR
  VAR lm AT %MW0 : ARRAY [1..2, -1..1] OF INT; END_VAR
  VAR k AT %IB0 : SINT; END_VAR
  VAR
    q0 AT %QB0 : SINT;
    q1 AT %QB1 : USINT;
    q2 AT %QB2 : SINT;
    q3 AT %QB3 : SINT;
    q4 AT %QB4 : SINT;
    q5 AT %QB5 : SINT;
    q6 AT %QB6 : SINT;
    q7 AT %QB7 : SINT;
    q8 AT %QB8 : SINT;
    q9 AT %QB9 : SINT;
    q10 AT %QB10 : SINT;
    q11 AT %QB11 : SINT;
    q12 AT %QB12 : SINT;
    q13 AT %QB13 : SINT;
    q14 AT %QB14 : SINT;
    q15 AT %QB15 : SINT;
    q16 AT %QB16 : SINT;
    q17 AT %QB17 : SINT;
    q18 AT %QB18 : SINT;
    q19 AT %QB19 : SINT;
    q20 AT %QB20 : SINT;
    q21 AT %QB21 : SINT;
    q22 AT %QB22 : SINT;
  END_VAR
  q0 := DINT_TO_SINT(SUM(a));
  q1 := DINT_TO_USINT(SUM(b));
  q2 := DINT_TO_SINT(TWICE(a));
  FILL(m);
  q3 := INT_TO_SINT(m[1, -1]);
  q4 := INT_TO_SINT(m[2, 1]);
  q5 := DINT_TO_SINT(LOWER_BOUND(b, 1));
  q6 := DINT_TO_SINT(UPPER_BOUND(m, 2));
  q7 := cnt.COUNT(row);
  q8 := INT_TO_SINT(LEN(s));
  q9 := INT_TO_SINT(lim);
  sc(k := 2, v := c, f := f, t := st, p := pr);
  q11 := INT_TO_SINT(c[2]);
  q12 := INT_TO_SINT(f[2]);
  q13 := INT_TO_SINT(LEN(st));
  q14 := pr.a;
  CASE k OF
    N - 4: q15 := 10;
    2..W - 1: q15 := 20;
  ELSE
    q15 := 30;
  END_CASE;
  q16 := DINT_TO_SINT(SUM(aa[2]));
  q17 := DINT_TO_SINT(SUM(aa[k MOD 2 + 1]));
  q18 := DINT_TO_SINT(SUM(m[2]));
  q19 := DINT_TO_SINT(SUM(m[k MOD 2 + 1]));
  r3 := m[1];
  q20 := INT_TO_SINT(r3[1]);
  q21 := DINT_TO_SINT(ROWSUM(m, 1));
  lm[2] := r3;
  r4 := lm[2];
  q22 := INT_TO_SINT(r4[0]);
  q10 := DINT_TO_SINT(UPPER_BOUND(m, k));
END_PROGRAM

(* ---- flexio.st ---- *)
(* An ARRAY[*] as a FUNCTION's and a method's input and output (Ed.3
   6.5.3): the caller's array itself, not a copy, as Siemens passes an
   FC's structured parameters (docs/dependencies.md).
   SUM adds an ARRAY[*] input. TWICE passes its input on to SUM. FILL
   writes all but the last element of an ARRAY[*] output; the output's
   elements are set to their initial value, 0, as the call starts. INC
   reads one ARRAY[*] and writes another. PICK reads one element.
   Worked by hand, k %IB0 (1, 2, 3):
   x: 1..3, [1, 2, 3]: SUM(x) 6, %QB0 6.
   y: 0..4, [9, 9, 9, 9, 9]. %QB1 := SUM(a := y), before FILL: 45 at
   tick 0. FILL(v := k, a => y) then makes y [k, k, k, k, 0]: %QB2 :=
   y[4] is 0 (it was 9: the output started from its initial value),
   %QB3 := y[0] is k: 1, 2, 3. So %QB1 is 4 at tick 1 and 8 at tick 2.
   TWICE(x) 12, %QB4 12.
   INC(src := x, dst => z), z: 1..3: z [2, 3, 4], %QB5 := z[3] 4.
   KC, a CONSTANT array [7, 8]: SUM(KC) 15, %QB6 15.
   The method TOP gives the last element: top.TOP(x) 3, %QB7 3.
   In order, the output after the inputs: FILL(5, w), w: 1..3 [5, 5,
   0]: %QB8 := w[1] 5, %QB9 := w[3] 0.
   A row of an array of arrays, aa [[1, 2, 3], [4, 5, 6]]: SUM(aa[2])
   15, %QB10 15.
   %QB11 := PICK(x, k + 1): x[2] 2, x[3] 3; at tick 2, x[4] is outside
   1..3, a fault (index), the statement stopped and %QB11 kept 3.
   reference-skip: ARRAY[*], LOWER_BOUND and UPPER_BOUND are Ed.3's, and
   CLASS; the reference compiler (Ed.2) has none. *)
FUNCTION SUM : DINT
  VAR_INPUT a : ARRAY [*] OF INT; END_VAR
  VAR i : DINT; END_VAR
  FOR i := LOWER_BOUND(a, 1) TO UPPER_BOUND(a, 1) DO
    SUM := SUM + a[i];
  END_FOR;
END_FUNCTION
FUNCTION TWICE : DINT
  VAR_INPUT a : ARRAY [*] OF INT; END_VAR
  TWICE := 2 * SUM(a);
END_FUNCTION
FUNCTION FILL
  VAR_INPUT v : INT; END_VAR
  VAR_OUTPUT a : ARRAY [*] OF INT; END_VAR
  VAR i : DINT; END_VAR
  FOR i := LOWER_BOUND(a, 1) TO UPPER_BOUND(a, 1) - 1 DO
    a[i] := v;
  END_FOR;
END_FUNCTION
FUNCTION INC
  VAR_INPUT src : ARRAY [*] OF INT; END_VAR
  VAR_OUTPUT dst : ARRAY [*] OF INT; END_VAR
  VAR i : DINT; END_VAR
  FOR i := LOWER_BOUND(src, 1) TO UPPER_BOUND(src, 1) DO
    dst[i] := src[i] + 1;
  END_FOR;
END_FUNCTION
FUNCTION PICK : INT
  VAR_INPUT a : ARRAY [*] OF INT; i : INT; END_VAR
  PICK := a[i];
END_FUNCTION
CLASS LAST
  METHOD PUBLIC TOP : INT
    VAR_INPUT a : ARRAY [*] OF INT; END_VAR
    TOP := a[UPPER_BOUND(a, 1)];
  END_METHOD
END_CLASS
CONFIGURATION c
  RESOURCE r ON PLC
    TASK t(INTERVAL := T#10ms, PRIORITY := 1);
    PROGRAM p WITH t : main;
  END_RESOURCE
END_CONFIGURATION
PROGRAM main
  VAR CONSTANT KC : ARRAY [1..2] OF INT := [7, 8]; END_VAR
  VAR
    x : ARRAY [1..3] OF INT := [1, 2, 3];
    y : ARRAY [0..4] OF INT := [5(9)];
    z : ARRAY [1..3] OF INT;
    w : ARRAY [1..3] OF INT := [3(1)];
    aa : ARRAY [1..2] OF ARRAY [0..2] OF INT := [[1, 2, 3], [4, 5, 6]];
    top : LAST;
  END_VAR
  VAR k AT %IB0 : SINT; END_VAR
  VAR
    q0 AT %QB0 : SINT;
    q1 AT %QB1 : SINT;
    q2 AT %QB2 : SINT;
    q3 AT %QB3 : SINT;
    q4 AT %QB4 : SINT;
    q5 AT %QB5 : SINT;
    q6 AT %QB6 : SINT;
    q7 AT %QB7 : SINT;
    q8 AT %QB8 : SINT;
    q9 AT %QB9 : SINT;
    q10 AT %QB10 : SINT;
    q11 AT %QB11 : SINT;
  END_VAR
  q0 := DINT_TO_SINT(SUM(x));
  q1 := DINT_TO_SINT(SUM(a := y));
  FILL(v := k, a => y);
  q2 := INT_TO_SINT(y[4]);
  q3 := INT_TO_SINT(y[0]);
  q4 := DINT_TO_SINT(TWICE(x));
  INC(src := x, dst => z);
  q5 := INT_TO_SINT(z[3]);
  q6 := DINT_TO_SINT(SUM(KC));
  q7 := INT_TO_SINT(top.TOP(x));
  FILL(5, w);
  q8 := INT_TO_SINT(w[1]);
  q9 := INT_TO_SINT(w[3]);
  q10 := DINT_TO_SINT(SUM(aa[2]));
  q11 := INT_TO_SINT(PICK(x, k + 1));
END_PROGRAM

(* ---- fnparams.st ---- *)
(* A FUNCTION's and a method's inputs, outputs, in-outs and results of a
   STRING, array or structure type (Ed.3 6.6.1.2, 6.6.2): LABEL's STRING
   result and STRING[3] input, given 'abcd' (cut to 'abc', flagged
   STRING_LENGTH at the call, as a block's input) or left to its initial
   value 'n'; RAMP's array result, assigned and given to SUM3's array
   input; SHIFT's structure input and result, its structure and STRING
   outputs, and its STRING in-out, which it cuts at the fifth '+'; a
   method's STRING result through an INTERFACE, overridden (Ed.3
   6.6.5.5); WRAP's WSTRING input and result.
   Worked by hand, the inputs v %IB0, pick %IX1.0:
   tick 0, v 7: qlab 'abc7'; xs 7, 8, 9: qsum 24 + 6 = 30; SHIFT of p
   (1, 2) by its d 10: q (11, -8), was (1, 2), tag 'ok', trail '+' (qtl
   1); nm the ANIMAL: 'anim'; ws '<' 16#263A '>': qw 16#263A, qwl 3; qdef
   TRUE ('n1'). The flag of the call giving LABEL 'abcd', line 109, stays.
   Tick 1, v 42: qlab 'abc42'; qsum 129 + 6 = 135; q (21, -18), was 11;
   qtl 2.
   Tick 2, v 255, pick TRUE: qlab 'abc255'; qsum 768 + 6 = 774; q (31,
   -28), was 21; qtl 3; nm the DOG: 'dog' (DOG's NAME, not ANIMAL's).
   Tick 3, v 0: qlab 'abc0', its sixth byte still '5' (a STRING in the
   image is its characters and a 0, the rest left); qsum 9; q (41, -38),
   was 31; qtl 4.
   Tick 4: q (51, -48), was 41; trail '+++++' cut to '++++', qtl 4.
   reference-skip: a method, an INTERFACE and WSTRING are Ed.3's; the
   reference compiler (Ed.2) has none. *)
TYPE PT :
  STRUCT
    x : INT;
    y : INT;
  END_STRUCT;
END_TYPE

FUNCTION LABEL : STRING[6]
  VAR_INPUT name : STRING[3] := 'n'; v : INT; END_VAR
  LABEL := CONCAT(name, INT_TO_STRING(v));
END_FUNCTION

FUNCTION SUM3 : INT
  VAR_INPUT xs : ARRAY[1..3] OF INT; END_VAR
  SUM3 := xs[1] + xs[2] + xs[3];
END_FUNCTION

FUNCTION RAMP : ARRAY[1..3] OF INT
  VAR_INPUT start : INT; END_VAR
  RAMP[1] := start;
  RAMP[2] := start + 1;
  RAMP[3] := start + 2;
END_FUNCTION

FUNCTION SHIFT : PT
  VAR_INPUT p : PT; d : INT := 10; END_VAR
  VAR_OUTPUT was : PT; tag : STRING[2]; END_VAR
  VAR_IN_OUT trail : STRING[4]; END_VAR
  was := p;
  SHIFT.x := p.x + d;
  SHIFT.y := p.y - d;
  tag := 'ok';
  trail := CONCAT(trail, '+');
END_FUNCTION

INTERFACE NAMED
  METHOD NAME : STRING[5]
  END_METHOD
END_INTERFACE

CLASS ANIMAL IMPLEMENTS NAMED
  METHOD PUBLIC NAME : STRING[5]
    NAME := 'anim';
  END_METHOD
END_CLASS

CLASS DOG EXTENDS ANIMAL
  METHOD PUBLIC OVERRIDE NAME : STRING[5]
    NAME := 'dog';
  END_METHOD
END_CLASS

FUNCTION WRAP : WSTRING[4]
  VAR_INPUT w : WSTRING[2]; END_VAR
  WRAP := CONCAT("<", w, ">");
END_FUNCTION

PROGRAM main
  VAR
    v AT %IB0 : USINT;
    pick AT %IX1.0 : BOOL;
    qlab AT %QB0 : STRING[6];
    qsum AT %QW8 : INT;
    qx AT %QW10 : INT;
    qy AT %QW12 : INT;
    qwx AT %QW14 : INT;
    qtag AT %QB16 : STRING[2];
    qtl AT %QB19 : USINT;
    qname AT %QB20 : STRING[5];
    qw AT %QW26 : WCHAR;
    qwl AT %QB28 : USINT;
    qdef AT %QX29.0 : BOOL;
  END_VAR
  VAR
    p : PT := (x := 1, y := 2);
    q, w : PT;
    xs : ARRAY[1..3] OF INT;
    trail : STRING[4];
    t : STRING[2];
    a : ANIMAL;
    d : DOG;
    nm : NAMED;
    ws : WSTRING[4];
  END_VAR
  qlab := LABEL(name := 'abcd', v := USINT_TO_INT(v));
  xs := RAMP(start := USINT_TO_INT(v));
  qsum := SUM3(xs := xs) + SUM3(xs := RAMP(start := 1));
  q := SHIFT(p := p, was => w, tag => t, trail := trail);
  p := q;
  qx := q.x;
  qy := q.y;
  qwx := w.x;
  qtag := t;
  qtl := INT_TO_USINT(LEN(trail));
  IF pick THEN
    nm := d;
  ELSE
    nm := a;
  END_IF;
  qname := nm.NAME();
  ws := WRAP(w := "${263A}");
  qw := ws[2];
  qwl := INT_TO_USINT(LEN(ws));
  qdef := LABEL(v := 1) = 'n1';
END_PROGRAM

CONFIGURATION Plant
  RESOURCE r ON PLC
    TASK fast(INTERVAL := T#10ms, PRIORITY := 1);
    PROGRAM p WITH fast : main;
  END_RESOURCE
END_CONFIGURATION

(* ---- hieraddr.st ---- *)
(* Single-level bit addresses and hierarchical addresses (Ed.3 Table
   16, 6.5.5.2). %IX9 is bit 9 of the input area, byte 1 bit 1; %I3 byte
   0 bit 3. A hierarchical address is where the platform's iecf_address
   puts it (docs/c-output.md §4); the harness's folds the levels into a
   byte from 256, each a hex digit, a bit address's last its bit:
   %IW2.5.7.1 is byte 256 + 0x2571 % 1024 = 625, %IX1.1.4 byte 273 bit
   4, %QX1.2.3 byte 274 bit 3, %QW3.3 byte 307, %QW7.7 byte 375, %MW1.1
   byte 273, %MW1.2.3 byte 547. Each written one is read back into the
   flat outputs. %IX1.1 (b9), %IX0.3 (b3), %IX273.4 TRUE, %IW625 41.
   Worked by hand:

   tick 0: out := iw + 1, 42 (Q0 2a 00); flags: b9, b3 and %IX1.1.4,
   2#111 (Q2 07); p, a structure at %MW1.1, p.y 2 (Q4 02 00); the
   block's w at %M*, put at %MW1.2.3 by VAR_CONFIG, 1 (Q10 01 00); %QW3.3 := iw, read back 41
   (Q6 29 00); s, at %Q* completed by %QW7.7 in VAR_CONFIG, 1 (Q8 01
   00); hb at %QX1.2.3 := b9, read back 1 (Q12 01).
   tick 1: p.y 4, w 2, s 2.
   reference-skip: the reference compiler takes one level. *)
TYPE Pt : STRUCT x : INT; y : INT; END_STRUCT; END_TYPE
FUNCTION_BLOCK blk
  VAR w AT %M* : UINT; END_VAR
  VAR_OUTPUT o : UINT; END_VAR
  w := w + 1;
  o := w;
END_FUNCTION_BLOCK
PROGRAM main
  VAR b9 AT %IX9 : BOOL; b3 AT %I3 : BOOL; END_VAR
  VAR iw AT %IW2.5.7.1 : INT; hb AT %QX1.2.3 : BOOL; p AT %MW1.1 : Pt; END_VAR
  VAR f : blk; END_VAR
  VAR out AT %QW0 : INT; flags AT %QB2 : BYTE; o2 AT %QW4 : INT; o3 AT %QW6 : INT; o4 AT %QW8 : INT;
      o5 AT %QW10 : UINT; o6 AT %QB12 : USINT; END_VAR
  VAR s AT %Q* : INT; END_VAR
  out := iw + 1;
  hb := b9;
  flags := BOOL_TO_BYTE(b9) OR SHL(BOOL_TO_BYTE(b3), 1) OR SHL(BOOL_TO_BYTE(%IX1.1.4), 2);
  p.y := p.y + 2;
  f();
  o2 := p.y;
  %QW3.3 := INT_TO_WORD(iw);
  o3 := WORD_TO_INT(%QW3.3);
  s := s + 1;
  o4 := s;
  o5 := f.o;
  o6 := BOOL_TO_USINT(hb);
END_PROGRAM
CONFIGURATION c
  RESOURCE r ON PLC
    TASK t(INTERVAL := T#10ms, PRIORITY := 1);
    PROGRAM pp WITH t : main;
  END_RESOURCE
  VAR_CONFIG r.pp.s AT %QW7.7 : INT; r.pp.f.w AT %MW1.2.3 : UINT; END_VAR
END_CONFIGURATION

(* ---- holders.st ---- *)
(* A structure or an array that holds function block instances, as a
   value everywhere an instance is one (docs/dependencies.md): a block's
   and a FUNCTION's input, output, in-out and result, an ARRAY[*] of
   instances, and a PROGRAM's connections of an array, a structure and
   an instance.
   CNT adds inc to n at each call; its inc stays as last given.
   Worked by hand, k %IB0 1, 2, 3:
   a(inc := k): a.n 1, 3, 6. h.c := a; h.k := k; arr[2] := a.
   f(h := h, cs := arr, io := h2, ios := arr2, o => h3):
     sum := h.c.n + cs[2].n + h.k: 3, 8, 15 (%QB0);
     o.c(inc := 3), o kept in f: 3, 6, 9, copied to h3 (%QB1); o.k :=
     sum, h3.k 3, 8, 15 (%QB2);
     io.c() is h2.c: at tick 0 its inc is 1, n 1; FNH below then calls
     it with inc := 10, which stays: 21 at tick 1, 41 at tick 2 (%QB3);
     ios[1](inc := 2) is arr2[1]: 2, 4, 6 (%QB4).
   r := FNH(h := h, o => o2, io := h2, fx := arr2):
     FNH := h; FNH.c() adds h.c's inc, k, to a.n: 2, 5, 9 (%QB5); FNH.k
     := h.k + 1: 2, 3, 4 (%QB6);
     o is set up at each call: o.c(inc := 4) 4 (%QB7); o.k := h.c.n 1,
     3, 6 (%QB8);
     io.c(inc := 10) on h2.c: 11, 31, 51 (%QB9);
     fx[UPPER_BOUND(fx, 1)]() is arr2[2]: 1, 2, 3 (%QB10).
   Connections, made before the program runs and after it:
     pa := ga, [10, 20, 30]; oa := pa; oa[2] := oa[2] + k; oa => gb,
     read at the next tick: gb[2] 0, 21, 22 (%QB11);
     pc := gc, and the program calls gc itself after: pc.n 0, 1, 2
     (%QB12); oc(inc := 5) => gd, at the next tick 0, 5, 10 (%QB13);
     ph := gh, the program then sets gh.k := k: ph.k 0, 1, 2 (%QB14);
     oh := ph; oh.k := ph.k + 100; oh => gi, at the next tick 0, 100,
     101 (%QB15).
   reference-skip: the reference compiler has no instance in a
   structure (tried in CI on instvalues). *)
FUNCTION_BLOCK CNT
  VAR_INPUT inc : INT := 1; END_VAR
  VAR_OUTPUT n : INT; END_VAR
  n := n + inc;
END_FUNCTION_BLOCK
TYPE HOLD : STRUCT c : CNT; k : INT; END_STRUCT; END_TYPE
FUNCTION_BLOCK FBH
  VAR_INPUT h : HOLD; cs : ARRAY [1..2] OF CNT; END_VAR
  VAR_OUTPUT o : HOLD; sum : INT; END_VAR
  VAR_IN_OUT io : HOLD; ios : ARRAY [1..2] OF CNT; END_VAR
  sum := h.c.n + cs[2].n + h.k;
  o.c(inc := 3);
  o.k := sum;
  io.c();
  ios[1](inc := 2);
END_FUNCTION_BLOCK
FUNCTION FNH : HOLD
  VAR_INPUT h : HOLD; END_VAR
  VAR_OUTPUT o : HOLD; END_VAR
  VAR_IN_OUT io : HOLD; fx : ARRAY [*] OF CNT; END_VAR
  FNH := h;
  FNH.c();
  FNH.k := h.k + 1;
  o.c(inc := 4);
  o.k := h.c.n;
  io.c(inc := 10);
  fx[UPPER_BOUND(fx, 1)]();
END_FUNCTION
CONFIGURATION c
  VAR_GLOBAL
    ga : ARRAY [1..3] OF INT := [10, 20, 30];
    gb : ARRAY [1..3] OF INT;
    gh, gi : HOLD;
    gc, gd : CNT;
  END_VAR
  RESOURCE r ON PLC
    TASK t(INTERVAL := T#10ms, PRIORITY := 1);
    PROGRAM p WITH t : main(pa := ga, ph := gh, pc := gc, oa => gb, oh => gi, oc => gd);
  END_RESOURCE
END_CONFIGURATION
PROGRAM main
  VAR_INPUT pa : ARRAY [1..3] OF INT; ph : HOLD; pc : CNT; END_VAR
  VAR_OUTPUT oa : ARRAY [1..3] OF INT; oh : HOLD; oc : CNT; END_VAR
  VAR_EXTERNAL
    gb : ARRAY [1..3] OF INT;
    gh, gi : HOLD;
    gc, gd : CNT;
  END_VAR
  VAR
    a : CNT;
    h, h2, h3, r, o2 : HOLD;
    arr, arr2 : ARRAY [1..2] OF CNT;
    f : FBH;
  END_VAR
  VAR k AT %IB0 : SINT; END_VAR
  VAR
    q0 AT %QB0 : SINT;
    q1 AT %QB1 : SINT;
    q2 AT %QB2 : SINT;
    q3 AT %QB3 : SINT;
    q4 AT %QB4 : SINT;
    q5 AT %QB5 : SINT;
    q6 AT %QB6 : SINT;
    q7 AT %QB7 : SINT;
    q8 AT %QB8 : SINT;
    q9 AT %QB9 : SINT;
    q10 AT %QB10 : SINT;
    q11 AT %QB11 : SINT;
    q12 AT %QB12 : SINT;
    q13 AT %QB13 : SINT;
    q14 AT %QB14 : SINT;
    q15 AT %QB15 : SINT;
  END_VAR
  a(inc := k);
  h.c := a;
  h.k := k;
  arr[2] := a;
  f(h := h, cs := arr, io := h2, ios := arr2, o => h3);
  q0 := INT_TO_SINT(f.sum);
  q1 := INT_TO_SINT(h3.c.n);
  q2 := INT_TO_SINT(h3.k);
  q3 := INT_TO_SINT(h2.c.n);
  q4 := INT_TO_SINT(arr2[1].n);
  r := FNH(h := h, o => o2, io := h2, fx := arr2);
  q5 := INT_TO_SINT(r.c.n);
  q6 := INT_TO_SINT(r.k);
  q7 := INT_TO_SINT(o2.c.n);
  q8 := INT_TO_SINT(o2.k);
  q9 := INT_TO_SINT(h2.c.n);
  q10 := INT_TO_SINT(arr2[2].n);
  q11 := INT_TO_SINT(gb[2]);
  oa := pa;
  oa[2] := oa[2] + k;
  q12 := INT_TO_SINT(pc.n);
  gc();
  q13 := INT_TO_SINT(gd.n);
  oc(inc := 5);
  q14 := INT_TO_SINT(ph.k);
  gh.k := k;
  q15 := INT_TO_SINT(gi.k);
  oh := ph;
  oh.k := ph.k + 100;
END_PROGRAM

(* ---- implicit.st ---- *)
(* The implicit-externals extension (docs/extensions.md): a PROGRAM, a
   FUNCTION_BLOCK and a FUNCTION use the configuration's globals without
   declaring them VAR_EXTERNAL, a CONSTANT one too; a FUNCTION that
   writes one has effects, so x := total + bump(1) reads total first
   (Ed.3 7.3.2).
   Worked by hand: tick 0, vin 2: qx 0 + 3 = 3 (total read as 0, then
   bump makes it 1 and gives 1 * 3), total 1 + 2 = 3, qs 3, qt 3.
   Tick 1, vin 5: qx 3 + 12 = 15 (total 3, bump makes it 4, 4 * 3),
   total 4 + 5 = 9, qs 9, qt 9.
   reference-skip: an extension, which the reference compiler has not. *)
FUNCTION bump : INT
VAR_INPUT n : INT; END_VAR
total := total + n;
bump := total * k3;
END_FUNCTION

FUNCTION_BLOCK counter
VAR_OUTPUT seen : INT; END_VAR
seen := total;
END_FUNCTION_BLOCK

PROGRAM main
VAR
  vin AT %IW0 : INT;
  qx AT %QW0 : INT;
  qs AT %QW2 : INT;
  qt AT %QW4 : INT;
END_VAR
VAR
  c : counter;
END_VAR
qx := total + bump(1);
total := total + vin;
c();
qs := c.seen;
qt := total;
END_PROGRAM

CONFIGURATION Plant
  VAR_GLOBAL
    total : INT;
  END_VAR
  VAR_GLOBAL CONSTANT
    k3 : INT := 3;
  END_VAR
  RESOURCE r ON PLC
    TASK fast(INTERVAL := T#10ms, PRIORITY := 1);
    PROGRAM p WITH fast : main;
  END_RESOURCE
END_CONFIGURATION

(* ---- inherit.st ---- *)
(* Inheritance and dynamic binding (Ed.3 6.6.5.5 to 6.6.5.8, 6.6.7.2.7
   to 6.6.7.3; OO.md step B): 6.6.5.6's CIRCLE, whose CF calls THIS.PI()
   and so in a CIRCLE2 runs CIRCLE2's PI; LIGHT2ROOM with SUPER.DAYTIME()
   (6.6.5.7.3), behind a LIGHTROOM in-out, and a block extending it;
   Figure 21's SUPER() chain, BASE, DERIVED_1, DERIVED_2; a DERIVED_1
   given to a BASE in-out and referenced by a REF_TO BASE, its body run
   (6.6.7.2.9 rule 4), its added input keeping its value (OO.md D7); an
   ABSTRACT SHAPE as a FUNCTION's in-out; a method called through a NULL
   reference (D8).
   Worked by hand, the inputs go %IX0.0 and night %IX0.1:
   tick 0, go FALSE, night FALSE: qa 300 (CIRCLE, PI 3.0), qb 314
   (CIRCLE2, PI 3.14), qr 30 (rr is c1); room1 day: LIGHT FALSE; room2
   day: LIGHT FALSE, LIGHT2 TRUE, Both FALSE; fr night: LIGHT TRUE,
   LIGHT2 FALSE (q byte 6 16#14); d2: x 3*(2+1)+0 9, c 9/5 1; qu1 6 (bb:
   x 5+1), qu2 19 (d1: SUPER() x 6, then 3*6+b, b 1); rb is bb, a 0:
   qref 1; qarea 1.
   Tick 1, go TRUE: qr 31 (rr is c2, 31.4); d2 x 10, c 10/1 10; rb is
   d1, a 1: x 3*2+1, qref 7; qarea 4.
   Tick 2, night TRUE: rooms night, fr day: byte 6 16#23; d2 x 11, c 1;
   qref 3*3+1 10; qarea 9.
   Tick 3, go FALSE: qr 30; d2 x 12, c 12; rb is bb, qref 4; qarea 16;
   qnull 1, then rn^.CF() faults NULL at line 194: the statement and the
   rest of the tick not run.
   reference-skip: EXTENDS, OVERRIDE and SUPER are Ed.3's; the
   reference compiler (Ed.2) has none. *)
CLASS CIRCLE
  METHOD PUBLIC PI : REAL
    PI := 3.0;
  END_METHOD
  METHOD PUBLIC CF : REAL
    VAR_INPUT d : REAL; END_VAR
    CF := THIS.PI() * d;
  END_METHOD
END_CLASS

CLASS CIRCLE2 EXTENDS CIRCLE
  METHOD PUBLIC OVERRIDE PI : REAL
    PI := 3.14;
  END_METHOD
END_CLASS

CLASS LIGHTROOM
  VAR PUBLIC LIGHT : BOOL; END_VAR
  METHOD PUBLIC DAYTIME
    LIGHT := FALSE;
  END_METHOD
  METHOD PUBLIC NIGHTTIME
    LIGHT := TRUE;
  END_METHOD
END_CLASS

CLASS LIGHT2ROOM EXTENDS LIGHTROOM
  VAR PUBLIC LIGHT2 : BOOL; END_VAR
  METHOD PUBLIC OVERRIDE DAYTIME
    SUPER.DAYTIME();
    LIGHT2 := TRUE;
  END_METHOD
  METHOD PUBLIC OVERRIDE NIGHTTIME
    SUPER.NIGHTTIME();
    LIGHT2 := FALSE;
  END_METHOD
  METHOD PUBLIC Both : BOOL
    Both := LIGHT AND LIGHT2;
  END_METHOD
END_CLASS

FUNCTION_BLOCK ROOM_CTRL
  VAR_INPUT night : BOOL; END_VAR
  VAR_IN_OUT RM : LIGHTROOM; END_VAR
  IF night THEN
    RM.NIGHTTIME();
  ELSE
    RM.DAYTIME();
  END_IF;
END_FUNCTION_BLOCK

FUNCTION_BLOCK FB_ROOM EXTENDS LIGHT2ROOM
  VAR_INPUT night : BOOL; END_VAR
  IF night THEN
    THIS.NIGHTTIME();
  ELSE
    THIS.DAYTIME();
  END_IF;
END_FUNCTION_BLOCK

FUNCTION_BLOCK BASE
  VAR_INPUT a : INT; END_VAR
  VAR_OUTPUT x : INT; END_VAR
  x := a + 1;
END_FUNCTION_BLOCK

FUNCTION_BLOCK DERIVED_1 EXTENDS BASE
  VAR_INPUT b : INT; END_VAR
  SUPER();
  x := 3 * x + b;
END_FUNCTION_BLOCK

FUNCTION_BLOCK DERIVED_2 EXTENDS DERIVED_1
  VAR_IN_OUT c : INT; END_VAR
  SUPER();
  c := x / c;
END_FUNCTION_BLOCK

FUNCTION_BLOCK USE
  VAR_IN_OUT io : BASE; END_VAR
  VAR_OUTPUT y : INT; END_VAR
  io(a := 5);
  y := io.x;
END_FUNCTION_BLOCK

CLASS ABSTRACT SHAPE
  METHOD PUBLIC ABSTRACT AREA : REAL
  END_METHOD
END_CLASS

CLASS SQUARE EXTENDS SHAPE
  VAR PUBLIC side : REAL; END_VAR
  METHOD PUBLIC OVERRIDE AREA : REAL
    AREA := side * side;
  END_METHOD
END_CLASS

FUNCTION total : INT
  VAR_IN_OUT s : SHAPE; END_VAR
  total := REAL_TO_INT(s.AREA());
END_FUNCTION

PROGRAM main
  VAR
    go AT %IX0.0 : BOOL;
    night AT %IX0.1 : BOOL;
    qa AT %QW0 : INT;
    qb AT %QW2 : INT;
    qr AT %QW4 : INT;
    ql1 AT %QX6.0 : BOOL;
    ql2 AT %QX6.1 : BOOL;
    ql3 AT %QX6.2 : BOOL;
    ql4 AT %QX6.3 : BOOL;
    ql5 AT %QX6.4 : BOOL;
    ql6 AT %QX6.5 : BOOL;
    qx AT %QW8 : INT;
    qc AT %QW10 : INT;
    qu1 AT %QW12 : INT;
    qu2 AT %QW14 : INT;
    qref AT %QW16 : INT;
    qarea AT %QW18 : INT;
    qnull AT %QB20 : BYTE;
  END_VAR
  VAR
    c1 : CIRCLE;
    c2 : CIRCLE2;
    rr, rn : REF_TO CIRCLE;
    room1 : LIGHTROOM;
    room2 : LIGHT2ROOM;
    ctrl : ROOM_CTRL;
    fr : FB_ROOM;
    d2 : DERIVED_2;
    cv : INT := 5;
    bb : BASE;
    d1 : DERIVED_1;
    u : USE;
    rb : REF_TO BASE;
    sq : SQUARE;
    n : INT;
  END_VAR
  qa := REAL_TO_INT(c1.CF(d := 100.0));
  qb := REAL_TO_INT(c2.CF(d := 100.0));
  IF go THEN rr := REF(c2); ELSE rr := REF(c1); END_IF;
  qr := REAL_TO_INT(rr^.CF(d := 10.0));
  ctrl(night := night, RM := room1);
  ctrl(night := night, RM := room2);
  fr(night := NOT night);
  ql1 := room1.LIGHT;
  ql2 := room2.LIGHT;
  ql3 := room2.LIGHT2;
  ql4 := room2.Both();
  ql5 := fr.LIGHT;
  ql6 := fr.LIGHT2;
  d2(a := 2, b := n, c := cv);
  qx := d2.x;
  qc := cv;
  d1.b := 1;
  u(io := bb);
  qu1 := u.y;
  u(io := d1);
  qu2 := u.y;
  IF go THEN rb := REF(d1); ELSE rb := REF(bb); END_IF;
  rb^(a := n);
  qref := rb^.x;
  sq.side := INT_TO_REAL(n + 1);
  qarea := total(s := sq);
  IF n = 3 THEN
    qnull := 1;
    qr := REAL_TO_INT(rn^.CF(d := 1.0));
  END_IF;
  n := n + 1;
END_PROGRAM

CONFIGURATION Plant
  RESOURCE r ON PLC
    TASK fast(INTERVAL := T#10ms, PRIORITY := 1);
    PROGRAM p WITH fast : main;
  END_RESOURCE
END_CONFIGURATION

(* ---- initexpr.st ---- *)
(* A variable's initial value that names variables and calls functions
   (the initial-expressions extension, docs/extensions.md), worked out as
   the variable is set up, in the order declared. Worked by hand:
   globals first: base 5, scaled base * Twice(3) = 5 * 6 = 30, RETAIN
   kept base + 1 = 6. Twice(x): its own y := x + 1, then (y - 1) * 2.
   main: a base * 2 = 10; b a + Twice(4) = 18; arr [a, b, 7], arr[1]
   18; p (x := a * 2), x 20, y its type's 9; c (d := b - a): Cnt sets
   up its own first, d 3 and q d * 10 = 30, then d is given 8; tm (PT :=
   pt0), T#2s; rg a * 20 = 200 into INT(0..100), clamped to 100 and
   flagged CONVERSION at its line (56), the first flag; s 'v10', LEN 3;
   RETAIN r kept * 2 = 12; m r + 1 = 13; the VAR_TEMP t b + 1 = 19 at
   each run. Each tick: c() runs its VAR_TEMP t := q + d, then q := t
   (38, then 46); n := acc.Add(t), the method's k := total + n (20,
   then 39); r := r + 1 (13, 14).
   A warm restart before tick 2: r keeps 14, kept 6; m is r + 1 = 15;
   c, acc set up again (q 38, n 20 at tick 2), r 15.
   %QB0 a 10, %QB1 b 18, %QB2 arr[1] 18, %QB3 p.x 20, %QB4 p.y 9, %QB5
   c.q, %QB6 rg 100, %QB7 LEN(s) 3, %QB8 scaled 30, %QB9 kept 6, %QB10
   r, %QB11 m, %QB12 n, %QX13.0 tm.PT = T#2s.
   reference-skip: a variable in an initial value is not IEC 61131-3. *)
TYPE Pt : STRUCT x : INT; y : INT := 9; END_STRUCT; END_TYPE

FUNCTION Twice : INT
  VAR_INPUT x : INT; END_VAR
  VAR y : INT := x + 1; END_VAR
  Twice := (y - 1) * 2;
END_FUNCTION

FUNCTION_BLOCK Cnt
  VAR_INPUT d : INT := 3; END_VAR
  VAR_OUTPUT q : INT := d * 10; END_VAR
  VAR_TEMP t : INT := q + d; END_VAR
  q := t;
END_FUNCTION_BLOCK

CLASS Accum
  VAR total : INT := 1; END_VAR
  METHOD PUBLIC Add : INT
    VAR_INPUT n : INT; END_VAR
    VAR k : INT := total + n; END_VAR
    total := k;
    Add := k;
  END_METHOD
END_CLASS

PROGRAM main
  VAR_EXTERNAL base : INT; scaled : INT; kept : INT; END_VAR
  VAR
    a : INT := base * 2;
    b : INT := a + Twice(4);
    arr : ARRAY[0..2] OF INT := [a, b, 7];
    p : Pt := (x := a * 2);
    c : Cnt := (d := b - a);
    pt0 : TIME := T#2s;
    tm : TON := (PT := pt0);
    rg : INT(0..100) := a * 20;
    s : STRING[8] := CONCAT('v', INT_TO_STRING(a));
    acc : Accum;
    n : INT;
  END_VAR
  VAR RETAIN r : INT := kept * 2; END_VAR
  VAR m : INT := r + 1; END_VAR
  VAR_TEMP t : INT := b + 1; END_VAR
  VAR
    q0 AT %QB0 : SINT;
    q1 AT %QB1 : SINT;
    q2 AT %QB2 : SINT;
    q3 AT %QB3 : SINT;
    q4 AT %QB4 : SINT;
    q5 AT %QB5 : SINT;
    q6 AT %QB6 : SINT;
    q7 AT %QB7 : SINT;
    q8 AT %QB8 : SINT;
    q9 AT %QB9 : SINT;
    q10 AT %QB10 : SINT;
    q11 AT %QB11 : SINT;
    q12 AT %QB12 : SINT;
    b0 AT %QX13.0 : BOOL;
  END_VAR
  c();
  n := acc.Add(t);
  r := r + 1;
  q0 := INT_TO_SINT(a);
  q1 := INT_TO_SINT(b);
  q2 := INT_TO_SINT(arr[1]);
  q3 := INT_TO_SINT(p.x);
  q4 := INT_TO_SINT(p.y);
  q5 := INT_TO_SINT(c.q);
  q6 := INT_TO_SINT(rg);
  q7 := INT_TO_SINT(LEN(s));
  q8 := INT_TO_SINT(scaled);
  q9 := INT_TO_SINT(kept);
  q10 := INT_TO_SINT(r);
  q11 := INT_TO_SINT(m);
  q12 := INT_TO_SINT(n);
  b0 := tm.PT = T#2s;
END_PROGRAM

CONFIGURATION cf
  VAR_GLOBAL base : INT := 5; scaled : INT := base * Twice(3); END_VAR
  VAR_GLOBAL RETAIN kept : INT := base + 1; END_VAR
  RESOURCE r ON x
    TASK tk(INTERVAL := T#10ms, PRIORITY := 1);
    PROGRAM p WITH tk : main;
  END_RESOURCE
END_CONFIGURATION

(* ---- inoutconst.st ---- *)
(* CODESYS's VAR_IN_OUT CONSTANT (the in-out-constant extension,
   docs/extensions.md): passed by reference and not written by the POU,
   given any value of its type - a literal, a constant, an expression, a
   variable - and a STRING of any length, read whole whatever the length
   declared. In a FUNCTION by name and in order, in a FUNCTION_BLOCK.
   Worked by hand, w = %IW0 each tick (2, 12, -3), lim clamped into 0..10
   and flagged as an input of a subrange is:
   r1 = addk(7, 'ab', q, arr, 3) = 7 + 2 + (1 + 2) + (10 + 30) + 3 = 55;
   r2 = addk(2w, long, KP, arr, w) = 2w + 10 + 7 + 40 + lim(w):
        63, 91 (12 clamped to 10, flagged), 51 (-3 to 0, flagged);
   r3 = addk(K5, CONCAT(long, 'xyz'), q, arr, w + 9) = 5 + 13 + 3 + 40
        + lim(w + 9): 71 (11 to 10, flagged), 71 (21, flagged), 67;
   f(inc := w + 1, tag := long): total 3, 16, 14; n = LEN(tag) = 10, a
   STRING[2] given ten characters. The flag is tick 0's, r3's line: the
   first stays until the platform clears it, and the host does not.
   reference-skip: VAR_IN_OUT CONSTANT is not IEC 61131-3. *)
TYPE pt : STRUCT x : INT; y : INT; END_STRUCT; END_TYPE
TYPE small : INT (0..10); END_TYPE

FUNCTION addk : INT
VAR_IN_OUT CONSTANT
  k : INT;
  s : STRING[4];
  p : pt;
  a : ARRAY[0..2] OF INT;
  lim : small;
END_VAR
addk := k + LEN(s) + p.x + p.y + a[0] + a[2] + lim;
END_FUNCTION

FUNCTION_BLOCK acc
VAR_IN_OUT CONSTANT inc : INT; tag : STRING[2]; END_VAR
VAR_OUTPUT total : INT; n : INT; END_VAR
total := total + inc;
n := LEN(tag);
END_FUNCTION_BLOCK

PROGRAM main
VAR
  v AT %IW0 : INT;
  r1 AT %QW0 : INT;
  r2 AT %QW2 : INT;
  r3 AT %QW4 : INT;
  r4 AT %QW6 : INT;
  r5 AT %QW8 : INT;
END_VAR
VAR
  long : STRING[20] := 'abcdefghij';
  q : pt := (x := 1, y := 2);
  arr : ARRAY[0..2] OF INT := [10, 20, 30];
  f : acc;
  w : INT;
END_VAR
VAR CONSTANT K5 : INT := 5; KP : pt := (x := 3, y := 4); END_VAR
w := v;
r1 := addk(k := 7, s := 'ab', p := q, a := arr, lim := 3);
r2 := addk(k := w * 2, s := long, p := KP, a := arr, lim := w);
r3 := addk(K5, CONCAT(long, 'xyz'), q, arr, w + 9);
f(inc := w + 1, tag := long);
r4 := f.total;
r5 := f.n;
END_PROGRAM

CONFIGURATION plant
  RESOURCE cpu ON PLC
    TASK t (INTERVAL := T#10ms, PRIORITY := 1);
    PROGRAM p WITH t : main;
  END_RESOURCE
END_CONFIGURATION

(* ---- inoutcopy.st ---- *)
(* An in-out given a variable at an address or of a subrange (Ed.3
   6.6.1.6 rule 6): given a copy, read before the call and stored back
   after it as an output is - clamped into the subrange and flagged
   CONVERSION. Siemens passes an elementary in-out so, copied in and
   back. To a FUNCTION (bump) and a FUNCTION_BLOCK (dbl), an element by
   a computed index too.
   Worked by hand, qw, qf 0, s 3, a[1] 0, t 1 at the start:
   Tick 0: qw 5, k 5; s 7, k 12; a[1] 2, k 14; qf 1; t 3.
   Tick 1: qw 10, k 10; bump gives 11, k 21, s stored back clamped to 9,
   flag CONVERSION on line 48; a[1] 4, k 25; qf 3; t 7.
   Tick 2: qw 15, k 15; s 13 clamped to 9, k 28; a[1] 6, k 34; qf 7;
   t 15 clamped to 9; the flag stays tick 1's.
   reference-skip: the reference compiler's C for an array element given
   as an in-out does not compile ("assignment to expression with array
   type"). *)
TYPE small : INT (0..9); END_TYPE

FUNCTION bump : INT
VAR_IN_OUT v : INT; END_VAR
VAR_INPUT d : INT; END_VAR
v := v + d;
bump := v;
END_FUNCTION

FUNCTION_BLOCK dbl
VAR_IN_OUT v : INT; END_VAR
v := v * 2 + 1;
END_FUNCTION_BLOCK

PROGRAM main
VAR
  qw AT %QW0 : INT;
  qs AT %QW2 : INT;
  qa AT %QW4 : INT;
  qk AT %QW6 : INT;
  qf AT %QW8 : INT;
  qt AT %QW10 : INT;
END_VAR
VAR
  s : small := 3;
  a : ARRAY[0..2] OF small;
  i : INT := 1;
  t : small := 1;
  k : INT;
  d : dbl;
END_VAR
k := bump(v := qw, d := 5);
k := k + bump(v := s, d := 4);
k := k + bump(v := a[i], d := 2);
d(v := qf);
d(v := t);
qs := s;
qa := a[1];
qt := t;
qk := k;
END_PROGRAM

CONFIGURATION Plant
  RESOURCE r ON PLC
    TASK fast(INTERVAL := T#10ms, PRIORITY := 1);
    PROGRAM p WITH fast : main;
  END_RESOURCE
END_CONFIGURATION

(* ---- inoutdata.st ---- *)
(* An array or a structure at an address, or reached through a
   reference, given to an in-out, to an ARRAY[*] input, output or
   in-out, of a FUNCTION and of a FUNCTION_BLOCK. No C object of its
   type is there (the image is read byte by byte), so the call is given
   a copy, stored back as it returns (docs/dependencies.md).
   SUM adds an ARRAY[*] input's first and last element. INC adds 1 to
   the first element of its ARRAY[*], to f[3] and to p.y; the block BMP
   does the same. SET writes 5 to the last element of its ARRAY[*]
   output, the others their initial 0.
   m at %MW0, 3 INTs; lp at %MW6, a PT; g at %MW10, 2 by 3 INTs. rm
   refers to m, r to x. Worked by hand, k %IB0 1, 2, 3:
   m[1] := k; m[3] := 10. SUM(m) k + 10: 11, 12, 13 (%QB0).
   g[2, 1] := 3; g[2, 3] := 4: SUM(g[2]), a row at an address, 7 (%QB1).
   SUM(rm^), through a reference, k + 10 (%QB2).
   INC(m, x, lp): m[1] k + 1; x[3] + 1; lp.y + 1.
   INC(g[j], rm^, ps[2]), j 1: g[1, 1] 1; m[3] 11; ps[2].y + 1.
   INC(r^, m, lp): x[1] + 1; m[3] 12; lp.y + 1.
   SET(a => g[1]): g[1] is [0, 0, 5].
   b(a := m, f := x, p := lp): m[1] k + 2; x[3] + 1; lp.y + 1.
   b(a := g[j], f := rm^, p := ps[j]): g[1, 1] 1; m[3] 13; ps[1].y + 1.
   So x[1] 1, 2, 3 (%QB3); x[3] 2, 4, 6 (%QB4); ps[2].y 1, 2, 3 (%QB5);
   ps[1].y 1, 2, 3 (%QB6); and in %M: m [k + 2, 0, 13], lp.y 3, 6, 9,
   g [[1, 0, 5], [3, 0, 4]].
   reference-skip: ARRAY[*] is Ed.3's; the reference compiler (Ed.2)
   has none. *)
TYPE PT : STRUCT x, y : INT; END_STRUCT; END_TYPE
FUNCTION SUM : INT
  VAR_INPUT a : ARRAY [*] OF INT; END_VAR
  SUM := a[LOWER_BOUND(a, 1)] + a[UPPER_BOUND(a, 1)];
END_FUNCTION
FUNCTION INC
  VAR_IN_OUT a : ARRAY [*] OF INT; f : ARRAY [1..3] OF INT; p : PT; END_VAR
  a[LOWER_BOUND(a, 1)] := a[LOWER_BOUND(a, 1)] + 1;
  f[3] := f[3] + 1;
  p.y := p.y + 1;
END_FUNCTION
FUNCTION SET
  VAR_OUTPUT a : ARRAY [*] OF INT; END_VAR
  a[UPPER_BOUND(a, 1)] := 5;
END_FUNCTION
FUNCTION_BLOCK BMP
  VAR_IN_OUT a : ARRAY [*] OF INT; f : ARRAY [1..3] OF INT; p : PT; END_VAR
  a[LOWER_BOUND(a, 1)] := a[LOWER_BOUND(a, 1)] + 1;
  f[3] := f[3] + 1;
  p.y := p.y + 1;
END_FUNCTION_BLOCK
CONFIGURATION c
  RESOURCE r ON PLC
    TASK t(INTERVAL := T#10ms, PRIORITY := 1);
    PROGRAM p WITH t : main;
  END_RESOURCE
END_CONFIGURATION
PROGRAM main
  VAR
    m AT %MW0 : ARRAY [1..3] OF INT;
    lp AT %MW6 : PT;
    g AT %MW10 : ARRAY [1..2, 1..3] OF INT;
  END_VAR
  VAR
    x : ARRAY [1..3] OF INT;
    r, rm : REF_TO ARRAY [1..3] OF INT;
    ps : ARRAY [1..2] OF PT;
    b : BMP;
    j : INT := 1;
  END_VAR
  VAR k AT %IB0 : SINT; END_VAR
  VAR
    q0 AT %QB0 : SINT;
    q1 AT %QB1 : SINT;
    q2 AT %QB2 : SINT;
    q3 AT %QB3 : SINT;
    q4 AT %QB4 : SINT;
    q5 AT %QB5 : SINT;
    q6 AT %QB6 : SINT;
  END_VAR
  m[1] := k;
  m[3] := 10;
  q0 := INT_TO_SINT(SUM(m));
  g[2, 1] := 3;
  g[2, 3] := 4;
  q1 := INT_TO_SINT(SUM(g[2]));
  rm := REF(m);
  q2 := INT_TO_SINT(SUM(rm^));
  INC(m, x, lp);
  INC(g[j], rm^, ps[2]);
  r := REF(x);
  INC(r^, m, lp);
  SET(a => g[1]);
  b(a := m, f := x, p := lp);
  b(a := g[j], f := rm^, p := ps[j]);
  q3 := INT_TO_SINT(x[1]);
  q4 := INT_TO_SINT(x[3]);
  q5 := INT_TO_SINT(ps[2].y);
  q6 := INT_TO_SINT(ps[1].y);
END_PROGRAM

(* ---- inouteffects.st ---- *)
(* FUNCTIONs with effects in the index of a variable given to an
   in-out, of a FUNCTION and of a block: each made once, in order, the
   element found before the call (an index out of bounds stops the
   statement first, docs/dependencies.md); a variable at an address or
   of a subrange given a copy, stored back after the call. Worked by
   hand, each tick from j 0:

   fadd(s[finc(j)], 20): j 1, s[1] 0 + 20 = 20 (40 at tick 1; inside
   0..50, no flag). fadd(la[finc(j)], 3): j 2, la[2] (Q1) 3, then 6.
   f(io := la[finc(j)], p := a[finc(j)]): j 3, then 4; la[3] (Q2) 1,
   then 2; a[4].y 1, then 2. From j 0 again: fp(a[finc(j)]): j 1, a[1].x
   10, then 20. finc(b[finc(j)]): j 1 again from 0, b[1] 1, then 2.
   Q4 s[1], Q5 a[4].y, Q6 a[1].x, Q7 b[1]; Q0 and Q3 untouched.
   reference-skip: VAR_IN_OUT of a FUNCTION, as `fnorder`. *)
TYPE small : SINT(0..50); END_TYPE
TYPE pt : STRUCT x : INT; y : INT; END_STRUCT; END_TYPE
FUNCTION finc : INT
  VAR_IN_OUT x : INT; END_VAR
  x := x + 1;
  finc := x;
END_FUNCTION
FUNCTION fadd : SINT
  VAR_IN_OUT x : SINT; END_VAR
  VAR_INPUT d : SINT; END_VAR
  x := x + d;
  fadd := x;
END_FUNCTION
FUNCTION fp : INT
  VAR_IN_OUT p : pt; END_VAR
  p.x := p.x + 10;
  fp := p.x;
END_FUNCTION
FUNCTION_BLOCK fb
  VAR_IN_OUT io : SINT; p : pt; END_VAR
  io := io + 1;
  p.y := p.y + 1;
END_FUNCTION_BLOCK
PROGRAM main
  VAR j : INT; s : ARRAY [1..4] OF small; a : ARRAY [1..4] OF pt; b : ARRAY [1..4] OF INT; f : fb; r : INT; END_VAR
  VAR la AT %QB0 : ARRAY [1..4] OF SINT; END_VAR
  VAR q4 AT %QB4 : USINT; q5 AT %QB5 : USINT; q6 AT %QB6 : USINT; q7 AT %QB7 : USINT; END_VAR
  j := 0;
  r := SINT_TO_INT(fadd(s[finc(j)], 20));
  r := SINT_TO_INT(fadd(la[finc(j)], 3));
  f(io := la[finc(j)], p := a[finc(j)]);
  j := 0;
  r := fp(a[finc(j)]);
  j := 0;
  r := finc(b[finc(j)]);
  q4 := SINT_TO_USINT(s[1]);
  q5 := INT_TO_USINT(a[4].y);
  q6 := INT_TO_USINT(a[1].x);
  q7 := INT_TO_USINT(b[1]);
END_PROGRAM
CONFIGURATION c RESOURCE r ON PLC TASK t(INTERVAL := T#10ms, PRIORITY := 1); PROGRAM p WITH t : main; END_RESOURCE END_CONFIGURATION

(* ---- inoutmember.st ---- *)
(* An instance's input or PUBLIC variable given to an in-out (Ed.3
   6.6.1.4: an in-out takes a variable; an input may be set from outside,
   6.6.7.2.2): the field itself, as an assignment from outside sets it.
   Inc adds 1 to its in-out. Worked by hand, tick by tick:
   f.a and f.pub 1, 2: f's q = a * 10 + pub, 11 then 22 (%QB0);
   fs[i].a, i 1: 1, 2, fs[1].q 10 then 20 (%QB1); b.v (a CLASS's
   PUBLIC) 1, 2 (%QB2); tm.PT (TON's input) T#1s then T#2s: %QX3.0 TRUE
   at tick 0, %QX3.1 TRUE at tick 1. And outputs taken into them, as
   an assignment from outside sets them: g(q => f.k), Gen's q 5, f.k 5
   (%QB4); Two(o => b.w), 2 (%QB5); ENO => f.ok TRUE (%QX6.0);
   SPLIT_DATE(IN := D#2024-03-05, YEAR => f.y), 2024 (%QW8, 16#07E8).
   reference-skip: VAR PUBLIC and CLASS are Ed.3's; the reference
   compiler (Ed.2) has neither. *)
FUNCTION Inc : INT
  VAR_IN_OUT c : INT; END_VAR
  c := c + 1;
  Inc := c;
END_FUNCTION

FUNCTION IncT : INT
  VAR_IN_OUT c : TIME; END_VAR
  c := c + T#1s;
  IncT := 0;
END_FUNCTION

FUNCTION Two : INT
  VAR_OUTPUT o : INT; END_VAR
  o := 2;
  Two := 1;
END_FUNCTION

FUNCTION_BLOCK Gen
  VAR_OUTPUT q : INT; END_VAR
  q := 5;
END_FUNCTION_BLOCK

FUNCTION_BLOCK Acc
  VAR_INPUT a : INT; k : INT; ok : BOOL; y : UINT; END_VAR
  VAR_OUTPUT q : INT; END_VAR
  VAR PUBLIC pub : INT; END_VAR
  q := a * 10 + pub;
END_FUNCTION_BLOCK

CLASS Box
  VAR PUBLIC v : INT; w : INT; END_VAR
END_CLASS

PROGRAM main
  VAR
    f : Acc;
    fs : ARRAY[0..1] OF Acc;
    b : Box;
    tm : TON;
    g : Gen;
    n : INT;
    i : INT := 1;
  END_VAR
  VAR
    q0 AT %QB0 : SINT;
    q1 AT %QB1 : SINT;
    q2 AT %QB2 : SINT;
    t1 AT %QX3.0 : BOOL;
    t2 AT %QX3.1 : BOOL;
    q4 AT %QB4 : SINT;
    q5 AT %QB5 : SINT;
    e6 AT %QX6.0 : BOOL;
    q8 AT %QW8 : UINT;
  END_VAR
  n := Inc(f.a);
  n := Inc(f.pub);
  f();
  n := Inc(fs[i].a);
  fs[i]();
  n := Inc(b.v);
  n := IncT(tm.PT);
  q0 := INT_TO_SINT(f.q);
  q1 := INT_TO_SINT(fs[1].q);
  q2 := INT_TO_SINT(b.v);
  t1 := tm.PT = T#1s;
  t2 := tm.PT = T#2s;
  g(q => f.k);
  n := Two(o => b.w);
  n := Two(EN := TRUE, ENO => f.ok);
  SPLIT_DATE(IN := D#2024-03-05, YEAR => f.y);
  q4 := INT_TO_SINT(f.k);
  q5 := INT_TO_SINT(b.w);
  e6 := f.ok;
  q8 := f.y;
END_PROGRAM

CONFIGURATION c
  RESOURCE r ON x
    TASK t(INTERVAL := T#10ms, PRIORITY := 1);
    PROGRAM p WITH t : main;
  END_RESOURCE
END_CONFIGURATION

(* ---- instances.st ---- *)
(* Function block and class instances besides a POU's own variable
   (Ed.3 6.6.3.3, 6.6.5.3, Table 11 rows 5a-7b, Figure 8 d and e): an
   ARRAY OF TON with [2(PT := T#20ms)], called as ts[i](...); an array of
   the user's CNT, each with its own initial value (an input, an output,
   a PUBLIC variable), called through an index from the input image and
   faulting INDEX when it is out of bounds; an array of a CLASS, its
   methods called on an element and an INTERFACE given one; a STRUCT with
   a TOF field whose PT the type gives (Table 11 7a), called as
   c.cooling(...); a FUNCTION_BLOCK holding an array of CNT; global
   instances, one named by a block's VAR_EXTERNAL, an array named by the
   program's; KEEPER, which keeps a RETAIN count, in a RETAIN array and a
   plain one, and in a plain global, across a warm restart; a RETAIN
   structure, its plain part kept too.
   Worked by hand, the inputs go %IX0.0, idx %IB1, ticks of 10 ms; USER
   calls the CNT it is given, so cs[idx] counts twice a tick:
   tick 0, go FALSE, idx 1: qtemp 16#11 (rc.temp 1, c.temp 1); ks[0] and
   kp[0] read 0, then count 1; b idle, sum 0; gc[0] 4; accs 11 and 11,
   qacc 11; cs[1] 10 (inc 5), cs[2] 50 (its n given), cs[3] 0.
   Tick 1, go TRUE, idx 2: ts[1] starts; c.cooling Q TRUE (qcool); qtemp
   16#22; qkr qkp 1; b counts cs 2 and 3, sum 5, gk 1; gc 8; accs 12, 23;
   cs[2] 52.
   Tick 2, idx 3: qtemp 16#33; qkr qkp 2; sum 10, gk 2; gc 12; accs 13,
   36; cs[3] 2.
   Tick 3, idx 1: ts[1] Q TRUE (ET 20 ms), ts[2] just started, Q FALSE
   (its PT 20 ms, not 0); qtemp 16#44; qkr qkp 3; sum 15, gk 3; gc 16;
   accs 14, 50; cs[1] 12, its lim (15 and 17 held there).
   Tick 4, go FALSE, idx 2: ts both FALSE; c.cooling still TRUE, PT not
   passed since IN fell; qtemp 16#55; qkr qkp 4; sum 15, gk 3; gc 20;
   accs 15, 65; cs[2] 54.
   A warm restart before tick 5: everything set anew but ks (RETAIN),
   rc (RETAIN, rc.temp 5 kept), and the RETAIN count of kp[0] and gk.
   Tick 5, idx 3: qcool FALSE (c anew); qtemp 16#61 (rc.temp 6, c.temp
   1); qkr 5 (ks[0].total kept), qkp 0 (kp[0].total anew); sum 0, gk.total
   0; gc 4; accs 11, 11; cs[1] 0, cs[2] 50, cs[3] 2.
   Tick 6, go TRUE, idx 4: qcool TRUE; qtemp 16#72; qkr qkp 6 (kp[0]'s
   count was kept); b counts 2 and 3, sum 5, gk 4 (its count kept); gc 8;
   accs 12, 23; then cs[4] given to u faults INDEX at line 158, u not
   called, qc1..qc3 as at tick 5.
   reference-skip: an array of instances, a CLASS, an INTERFACE and a
   PUBLIC variable are Ed.3's; the reference compiler (Ed.2) has none. *)
FUNCTION_BLOCK CNT
  VAR_INPUT inc : INT := 1; END_VAR
  VAR_OUTPUT n : INT; END_VAR
  VAR PUBLIC lim : INT := 100; END_VAR
  n := n + inc;
  IF n > lim THEN
    n := lim;
  END_IF;
END_FUNCTION_BLOCK

FUNCTION_BLOCK KEEPER
  VAR_OUTPUT total : INT; END_VAR
  VAR RETAIN kept : INT; END_VAR
  kept := kept + 1;
  total := kept;
END_FUNCTION_BLOCK

INTERFACE SHOW
  METHOD GET : INT
  END_METHOD
END_INTERFACE

CLASS ACC IMPLEMENTS SHOW
  VAR PUBLIC v : INT; END_VAR
  METHOD PUBLIC ADD
    VAR_INPUT x : INT; END_VAR
    v := v + x;
  END_METHOD
  METHOD PUBLIC GET : INT
    GET := v;
  END_METHOD
END_CLASS

TYPE COOLER :
  STRUCT
    temp : INT;
    cooling : TOF := (PT := T#20ms);
  END_STRUCT;
END_TYPE

FUNCTION_BLOCK USER
  VAR_IN_OUT c : CNT; END_VAR
  c();
END_FUNCTION_BLOCK

FUNCTION_BLOCK BANK
  VAR_INPUT go : BOOL; END_VAR
  VAR_OUTPUT sum : INT; END_VAR
  VAR cs : ARRAY[0..1] OF CNT := [(inc := 2), (inc := 3)]; END_VAR
  VAR_EXTERNAL gk : KEEPER; END_VAR
  IF go THEN
    cs[0]();
    cs[1]();
    gk();
  END_IF;
  sum := cs[0].n + cs[1].n;
END_FUNCTION_BLOCK

PROGRAM main
  VAR
    go AT %IX0.0 : BOOL;
    idx AT %IB1 : USINT;
    qt1 AT %QX0.0 : BOOL;
    qt2 AT %QX0.1 : BOOL;
    qcool AT %QX0.2 : BOOL;
    qc1 AT %QW2 : INT;
    qc2 AT %QW4 : INT;
    qc3 AT %QW6 : INT;
    qacc AT %QW8 : INT;
    qbank AT %QW10 : INT;
    qkr AT %QW12 : INT;
    qkp AT %QW14 : INT;
    qg AT %QW16 : INT;
    qgc AT %QW18 : INT;
    qtemp AT %QW20 : INT;
  END_VAR
  VAR
    ts : ARRAY[1..2] OF TON := [2(PT := T#20ms)];
    cs : ARRAY[1..3] OF CNT := [(inc := 5, lim := 12), (n := 50)];
    accs : ARRAY[0..1] OF ACC := [(v := 10)];
    c : COOLER;
    b : BANK;
    s : SHOW;
    u : USER;
    kp : ARRAY[0..1] OF KEEPER;
  END_VAR
  VAR RETAIN
    ks : ARRAY[0..1] OF KEEPER;
    rc : COOLER;
  END_VAR
  VAR_EXTERNAL
    gk : KEEPER;
    gc : ARRAY[0..1] OF CNT;
  END_VAR
  ts[1](IN := go);
  ts[2](IN := ts[1].Q);
  qt1 := ts[1].Q;
  qt2 := ts[2].Q;
  c.cooling(IN := go);
  qcool := c.cooling.Q;
  c.temp := c.temp + 1;
  rc.temp := rc.temp + 1;
  qtemp := rc.temp * 16 + c.temp;
  qkr := ks[0].total;
  qkp := kp[0].total;
  ks[0]();
  kp[0]();
  b(go := go);
  qbank := b.sum;
  qg := gk.total;
  gc[0]();
  qgc := gc[0].n;
  (* An index the generator does not fold: checked, as idx is. *)
  accs[idx - idx].ADD(x := 1);
  accs[1].ADD(x := accs[0].v);
  s := accs[1];
  qacc := s.GET();
  u(c := cs[idx]);
  cs[idx]();
  qc1 := cs[1].n;
  qc2 := cs[2].n;
  qc3 := cs[3].n;
END_PROGRAM

CONFIGURATION Plant
  VAR_GLOBAL
    gk : KEEPER;
    gc : ARRAY[0..1] OF CNT := [(inc := 4)];
  END_VAR
  RESOURCE r ON PLC
    TASK fast(INTERVAL := T#10ms, PRIORITY := 1);
    PROGRAM p WITH fast : main;
  END_RESOURCE
END_CONFIGURATION

(* ---- instvalues.st ---- *)
(* Function block instances as values (Ed.3 Table 72 1d, Table 42 9a,
   6.6.1.4 rule 4; docs/dependencies.md): an instance assigned is copied
   whole, every variable of it; one given as an input is a copy, read
   in the POU it is given to.
   CNT adds inc to n at each call. Worked by hand, k %IB0 1, 2, 3:
   a(inc := k): a.n 1, 3, 6.
   b := a; b(): b has a's n and inc, then adds: 2, 5, 9 (%QB0); a is as
   it was: 1, 3, 6 (%QB1).
   h.c := a; h2 := h, a structure holding an instance; h2.c() adds k:
   h2.c.n 2, 5, 9 (%QB2); h.c.n 1, 3, 6 (%QB3).
   arr[1] := a; arr2 := arr, an array of instances: arr2[1].n 1, 3, 6
   (%QB4); arr2[2].n 0 (%QB5).
   PEEK takes a CNT as an input and gives n * 10 + inc: PEEK(a) 11, 32,
   63 (%QB6); PEEK() has the instance's initial values, n 0, inc 1: 1
   (%QB7).
   WATCH takes a CNT as an input, c, and has one as an output, own,
   which it calls with inc := 5. w(c := a, own => d): seen := c.n, 1,
   3, 6 (%QB8); d is a copy of own: d.n 5, 10, 15 (%QB9); the copy kept
   in w, w.c.inc, is k: 1, 2, 3 (%QB10).
   A standard block: t1(IN := TRUE, PT := T#15ms), ticks 10 ms apart:
   ET 0, 10, 20 ms, so Q at tick 2; t2 := t1 has it: %QX11.0 0, 0, 1.
   An input set apart from a call: w.c := b; w.c.n 2, 5, 9 (%QB12).
   A FUNCTION's result an instance: MAKE(amt) sets its result's inc and
   calls it once; e := MAKE(k): e.n 1, 2, 3 (%QB13).
   A FUNCTION's own instance and its output one keep nothing from call
   to call: WORK calls c twice with inc 4, c.n 8, its result (%QB14),
   and o once with inc 7; WORK(o => f): f.n 7 at every tick (%QB15).
   reference-skip: the reference compiler refuses an instance in a
   structure, as a FUNCTION's result and as a FUNCTION's variable. *)
FUNCTION_BLOCK CNT
  VAR_INPUT inc : INT := 1; END_VAR
  VAR_OUTPUT n : INT; END_VAR
  n := n + inc;
END_FUNCTION_BLOCK
TYPE HOLD : STRUCT c : CNT; k : INT; END_STRUCT; END_TYPE
FUNCTION PEEK : INT
  VAR_INPUT c : CNT; END_VAR
  PEEK := c.n * 10 + c.inc;
END_FUNCTION
FUNCTION MAKE : CNT
  VAR_INPUT amt : INT; END_VAR
  MAKE.inc := amt;
  MAKE();
END_FUNCTION
FUNCTION WORK : INT
  VAR c : CNT; END_VAR
  VAR_OUTPUT o : CNT; END_VAR
  c(inc := 4);
  c();
  o(inc := 7);
  WORK := c.n;
END_FUNCTION
FUNCTION_BLOCK WATCH
  VAR_INPUT c : CNT; END_VAR
  VAR_OUTPUT seen : INT; own : CNT; END_VAR
  seen := c.n;
  own(inc := 5);
END_FUNCTION_BLOCK
CONFIGURATION c
  RESOURCE r ON PLC
    TASK t(INTERVAL := T#10ms, PRIORITY := 1);
    PROGRAM p WITH t : main;
  END_RESOURCE
END_CONFIGURATION
PROGRAM main
  VAR
    a, b, d, e, f : CNT;
    h, h2 : HOLD;
    arr, arr2 : ARRAY [1..2] OF CNT;
    w : WATCH;
    t1, t2 : TON;
  END_VAR
  VAR k AT %IB0 : SINT; END_VAR
  VAR
    q0 AT %QB0 : SINT;
    q1 AT %QB1 : SINT;
    q2 AT %QB2 : SINT;
    q3 AT %QB3 : SINT;
    q4 AT %QB4 : SINT;
    q5 AT %QB5 : SINT;
    q6 AT %QB6 : SINT;
    q7 AT %QB7 : SINT;
    q8 AT %QB8 : SINT;
    q9 AT %QB9 : SINT;
    q10 AT %QB10 : SINT;
    q11 AT %QX11.0 : BOOL;
    q12 AT %QB12 : SINT;
    q13 AT %QB13 : SINT;
    q14 AT %QB14 : SINT;
    q15 AT %QB15 : SINT;
  END_VAR
  a(inc := k);
  b := a;
  b();
  q0 := INT_TO_SINT(b.n);
  q1 := INT_TO_SINT(a.n);
  h.c := a;
  h2 := h;
  h2.c();
  q2 := INT_TO_SINT(h2.c.n);
  q3 := INT_TO_SINT(h.c.n);
  arr[1] := a;
  arr2 := arr;
  q4 := INT_TO_SINT(arr2[1].n);
  q5 := INT_TO_SINT(arr2[2].n);
  q6 := INT_TO_SINT(PEEK(a));
  q7 := INT_TO_SINT(PEEK());
  w(c := a, own => d);
  q8 := INT_TO_SINT(w.seen);
  q9 := INT_TO_SINT(d.n);
  q10 := INT_TO_SINT(w.c.inc);
  t1(IN := TRUE, PT := T#15ms);
  t2 := t1;
  q11 := t2.Q;
  w.c := b;
  q12 := INT_TO_SINT(w.c.n);
  e := MAKE(k);
  q13 := INT_TO_SINT(e.n);
  q14 := INT_TO_SINT(WORK(o => f));
  q15 := INT_TO_SINT(f.n);
END_PROGRAM

(* ---- interfaces.st ---- *)
(* Interfaces (Ed.3 6.6.6; OO.md step C): 6.6.6.5.3's ROOM and its
   ROOM_CTRL, which takes any ROOM as an input: a LIGHTROOM, a
   LIGHT2ROOM through THIS in a method of its base (its own overrides
   run), a FullT whose ABSTRACT base HALF implements DAYTIME only, a
   DIMMER of DIMMED, an interface extending ROOM; one ROOM holding a
   DIMMER or a LIGHT2ROOM, and ?= from it to a DIMMED and to a REF_TO
   DIMMER (6.6.6.7), NULL when it holds the other; ?= from a REF_TO
   LIGHTROOM to a REF_TO LIGHT2ROOM; = of interfaces; a FUNCTION taking a
   DIMMED, a ROOM of its own given it; a method with an output and ENO
   through its interface; a method called through a NULL interface
   (OO.md D8).
   Worked by hand, the inputs night %IX0.0, pick %IX0.1, stop %IX0.2,
   pct %IB1:
   tick 0, all FALSE, pct 0: room1 day: LIGHT FALSE; room2 through THIS
   night: LIGHT TRUE, LIGHT2 FALSE; full day: day TRUE (HALF's); dm day:
   lvl 0; r is room2, so d ?= r NULL (qnull), rd ?= r NULL; qof -1 (the
   FUNCTION's ROOM NULL); qx 0; qsame FALSE; rl is room1, rl2 ?= rl NULL;
   qcalls 4. Q byte 0: 16#1A.
   Tick 1, night TRUE, pick TRUE, pct 30: room1 night LIGHT TRUE; room2
   day: LIGHT FALSE, LIGHT2 TRUE; full night: day FALSE (FullT's); dm
   night lvl 100; r is dm: d and rd it; qof 30 (LEVEL 30); qx 80 (LEVEL
   80, not clipped); qsame TRUE; rl is room2, rl2 it; qlvl 80; qcalls 8.
   Q byte 0: 16#E5.
   Tick 2, pct 80: as tick 1, qof 80, then LEVEL 130 clipped: lvl 100,
   qx 100, qclip TRUE; qcalls 12.
   Tick 3, night FALSE, pick FALSE, stop TRUE: as tick 0, qcalls 16;
   then none.DAYTIME() faults NULL at line 200, the call not made.
   reference-skip: INTERFACE, IMPLEMENTS and ?= are Ed.3's; the
   reference compiler (Ed.2) has none. *)
INTERFACE ROOM
  METHOD DAYTIME
  END_METHOD
  METHOD NIGHTTIME
  END_METHOD
END_INTERFACE

INTERFACE DIMMED EXTENDS ROOM
  METHOD LEVEL : INT
    VAR_INPUT pct : INT; END_VAR
    VAR_OUTPUT clipped : BOOL; END_VAR
  END_METHOD
END_INTERFACE

FUNCTION_BLOCK ROOM_CTRL
  VAR_INPUT RM : ROOM; night : BOOL; END_VAR
  VAR_OUTPUT calls : INT; END_VAR
  IF RM = NULL THEN
    RETURN;
  END_IF;
  IF night THEN
    RM.NIGHTTIME();
  ELSE
    RM.DAYTIME();
  END_IF;
  calls := calls + 1;
END_FUNCTION_BLOCK

CLASS LIGHTROOM IMPLEMENTS ROOM
  VAR PUBLIC LIGHT : BOOL; END_VAR
  METHOD PUBLIC DAYTIME
    LIGHT := FALSE;
  END_METHOD
  METHOD PUBLIC NIGHTTIME
    LIGHT := TRUE;
  END_METHOD
  METHOD PUBLIC SELF_CTRL
    VAR_IN_OUT c : ROOM_CTRL; END_VAR
    VAR_INPUT n : BOOL; END_VAR
    c(RM := THIS, night := n);
  END_METHOD
END_CLASS

CLASS LIGHT2ROOM EXTENDS LIGHTROOM
  VAR PUBLIC LIGHT2 : BOOL; END_VAR
  METHOD PUBLIC OVERRIDE DAYTIME
    SUPER.DAYTIME();
    LIGHT2 := TRUE;
  END_METHOD
  METHOD PUBLIC OVERRIDE NIGHTTIME
    SUPER.NIGHTTIME();
    LIGHT2 := FALSE;
  END_METHOD
END_CLASS

CLASS DIMMER IMPLEMENTS DIMMED
  VAR PUBLIC lvl : INT; END_VAR
  METHOD PUBLIC DAYTIME
    lvl := 0;
  END_METHOD
  METHOD PUBLIC NIGHTTIME
    lvl := 100;
  END_METHOD
  METHOD PUBLIC LEVEL : INT
    VAR_INPUT pct : INT; END_VAR
    VAR_OUTPUT clipped : BOOL; END_VAR
    clipped := pct > 100;
    ENO := NOT clipped;
    IF clipped THEN
      lvl := 100;
    ELSE
      lvl := pct;
    END_IF;
    LEVEL := lvl;
  END_METHOD
END_CLASS

FUNCTION_BLOCK ABSTRACT HALF IMPLEMENTS ROOM
  VAR_OUTPUT day : BOOL; END_VAR
  METHOD PUBLIC DAYTIME
    day := TRUE;
  END_METHOD
END_FUNCTION_BLOCK

FUNCTION_BLOCK FullT EXTENDS HALF
  METHOD PUBLIC NIGHTTIME
    day := FALSE;
  END_METHOD
END_FUNCTION_BLOCK

FUNCTION LEVEL_OF : INT
  VAR_INPUT d : DIMMED; pct : INT; END_VAR
  VAR r : ROOM; END_VAR
  r := d;
  IF r = NULL THEN
    LEVEL_OF := -1;
    RETURN;
  END_IF;
  LEVEL_OF := d.LEVEL(pct := pct);
END_FUNCTION

PROGRAM main
  VAR
    night AT %IX0.0 : BOOL;
    pick AT %IX0.1 : BOOL;
    stop AT %IX0.2 : BOOL;
    pct AT %IB1 : USINT;
    ql1 AT %QX0.0 : BOOL;
    ql2 AT %QX0.1 : BOOL;
    ql3 AT %QX0.2 : BOOL;
    qday AT %QX0.3 : BOOL;
    qnull AT %QX0.4 : BOOL;
    qrd AT %QX0.5 : BOOL;
    qsame AT %QX0.6 : BOOL;
    qdown AT %QX0.7 : BOOL;
    qlvl AT %QW2 : INT;
    qof AT %QW4 : INT;
    qx AT %QW6 : INT;
    qclip AT %QX8.0 : BOOL;
    qcalls AT %QW10 : INT;
  END_VAR
  VAR
    room1 : LIGHTROOM;
    room2 : LIGHT2ROOM;
    dm : DIMMER;
    full : FullT;
    ctrl : ROOM_CTRL;
    r : ROOM;
    d : DIMMED;
    none : ROOM;
    rd : REF_TO DIMMER;
    rl : REF_TO LIGHTROOM;
    rl2 : REF_TO LIGHT2ROOM;
    cl : BOOL;
  END_VAR
  ctrl(RM := room1, night := night);
  room2.SELF_CTRL(c := ctrl, n := NOT night);
  ctrl(RM := full, night := night);
  ctrl(RM := dm, night := night);
  IF pick THEN
    r := dm;
  ELSE
    r := room2;
  END_IF;
  d ?= r;
  qnull := d = NULL;
  rd ?= r;
  qrd := rd <> NULL;
  qof := LEVEL_OF(d := d, pct := pct);
  qx := 0;
  qclip := FALSE;
  IF d <> NULL THEN
    qx := d.LEVEL(pct := USINT_TO_INT(pct) + 50, clipped => cl);
    qclip := cl;
  END_IF;
  qsame := r = d;
  IF night THEN
    rl := REF(room2);
  ELSE
    rl := REF(room1);
  END_IF;
  rl2 ?= rl;
  qdown := rl2 <> NULL;
  ql1 := room1.LIGHT;
  ql2 := room2.LIGHT;
  ql3 := room2.LIGHT2;
  qday := full.day;
  qlvl := dm.lvl;
  qcalls := ctrl.calls;
  IF stop THEN
    none.DAYTIME();
  END_IF;
END_PROGRAM

CONFIGURATION Plant
  RESOURCE r ON PLC
    TASK fast(INTERVAL := T#10ms, PRIORITY := 1);
    PROGRAM p WITH fast : main;
  END_RESOURCE
END_CONFIGURATION

(* ---- itfplaces.st ---- *)
(* Interfaces wherever a variable can be (Ed.3 6.6.6.5.1: "This rule
   applies for all cases where variables may be used"): array elements
   and structure fields, a VAR_GLOBAL, initial values that are instances
   (a local's, a global's), a FUNCTION's result, output and input with an
   initial value, a block's output (taken into an element and read from
   outside), a method's result and output, a method through an
   interface's table giving an interface, ?= into an element, = of
   elements, an element's method called, NULL there faulting (OO.md D8).
   Worked by hand, k %IB0 and stop %IX1.0; ID_OF gives a ROOM's id, 0
   for NULL; l1 is 1, gl 2, dm 3:
   tick 0, k 0: arr [l1, dm, l1] (arr[0] := l1 after dm; arr[2] the
   block's output, h.r = l1); hs[1].r = g = gl; SWAP's b not given, so
   hs[2].r NULL and tmp l1; d ?= arr[1] dm; darr[1] ?= arr[0] NULL.
   qa..qi 1 3 1 2 0 1 3 0 1; tmp := darr[0].ME() dm: qj 3; dm.GIVE puts
   dm in hs[2].r: qk 3; ql LEVEL(0) 0; arr[0] = arr[1] FALSE, hs[1].r =
   rg TRUE, darr[1] = NULL TRUE: Q byte 0 16#06.
   Tick 1, k 1: arr [dm, l1, l1]; tmp dm; d ?= l1 NULL; darr[1] ?= dm.
   qa..qi 3 1 1 2 0 3 0 3 1, qj 3, qk 3, ql 10; byte 0 16#02.
   Tick 2, k 2: arr [dm, dm, l1]; d dm, darr[1] dm. qa..qi 3 3 1 2 0 3 3
   3 1, qj 3, qk 3, ql 20; byte 0 16#03.
   Tick 3, stop TRUE: as tick 2, then hs[2].r NULL, its DAYTIME() faults
   NULL, the call not made.
   reference-skip: INTERFACE and CLASS are Ed.3's; the reference
   compiler (Ed.2) has neither. *)
INTERFACE ROOM
  METHOD DAYTIME
  END_METHOD
  METHOD NAME : SINT
  END_METHOD
END_INTERFACE

INTERFACE DIMMED EXTENDS ROOM
  METHOD LEVEL : INT
    VAR_INPUT pct : INT; END_VAR
  END_METHOD
  METHOD ME : DIMMED
  END_METHOD
END_INTERFACE

CLASS LIGHTROOM IMPLEMENTS ROOM
  VAR PUBLIC id : SINT; LIGHT : BOOL; END_VAR
  METHOD PUBLIC DAYTIME
    LIGHT := NOT LIGHT;
  END_METHOD
  METHOD PUBLIC NAME : SINT
    NAME := id;
  END_METHOD
END_CLASS

CLASS DIMMER IMPLEMENTS DIMMED
  VAR PUBLIC id : SINT; lvl : INT; END_VAR
  METHOD PUBLIC DAYTIME
    lvl := 0;
  END_METHOD
  METHOD PUBLIC NAME : SINT
    NAME := id;
  END_METHOD
  METHOD PUBLIC LEVEL : INT
    VAR_INPUT pct : INT; END_VAR
    lvl := pct;
    LEVEL := lvl;
  END_METHOD
  METHOD PUBLIC ME : DIMMED
    ME := THIS;
  END_METHOD
  METHOD PUBLIC GIVE
    VAR_OUTPUT r : ROOM; END_VAR
    r := THIS;
  END_METHOD
END_CLASS

TYPE HOLDER : STRUCT
  r : ROOM;
  n : INT;
END_STRUCT;
END_TYPE

FUNCTION_BLOCK PICKER
  VAR_INPUT a : ROOM; END_VAR
  VAR_OUTPUT o : ROOM; END_VAR
  o := a;
END_FUNCTION_BLOCK

FUNCTION PICK : ROOM
  VAR_INPUT a : ROOM; END_VAR
  PICK := a;
END_FUNCTION

FUNCTION SWAP
  VAR_INPUT a : ROOM; b : ROOM := NULL; END_VAR
  VAR_OUTPUT x : ROOM; y : ROOM; END_VAR
  x := b;
  y := a;
END_FUNCTION

FUNCTION ID_OF : SINT
  VAR_INPUT r : ROOM; END_VAR
  IF r = NULL THEN
    ID_OF := 0;
  ELSE
    ID_OF := r.NAME();
  END_IF;
END_FUNCTION

CONFIGURATION plant
  VAR_GLOBAL
    gl : LIGHTROOM := (id := 2);
    g : ROOM := gl;
  END_VAR
  RESOURCE cpu ON PLC
    TASK fast(INTERVAL := T#10ms, PRIORITY := 1);
    PROGRAM p WITH fast : main;
  END_RESOURCE
END_CONFIGURATION

PROGRAM main
  VAR_EXTERNAL
    g : ROOM;
    gl : LIGHTROOM;
  END_VAR
  VAR
    l1 : LIGHTROOM := (id := 1);
    dm : DIMMER := (id := 3);
    arr : ARRAY[0..2] OF ROOM;
    darr : ARRAY[0..1] OF DIMMED := [dm, NULL];
    h : HOLDER := (r := l1, n := 3);
    hs : ARRAY[1..2] OF HOLDER;
    pk : PICKER;
    i : INT;
    d : DIMMED;
    tmp : ROOM;
    rg : ROOM := gl;
  END_VAR
  VAR
    k AT %IB0 : USINT;
    stop AT %IX1.0 : BOOL;
    qx0 AT %QX0.0 : BOOL;
    qx1 AT %QX0.1 : BOOL;
    qx2 AT %QX0.2 : BOOL;
    qa AT %QB1 : SINT;
    qb AT %QB2 : SINT;
    qc AT %QB3 : SINT;
    qd AT %QB4 : SINT;
    qe AT %QB5 : SINT;
    qf AT %QB6 : SINT;
    qg AT %QB7 : SINT;
    qh AT %QB8 : SINT;
    qi AT %QB9 : SINT;
    qj AT %QB10 : SINT;
    qk AT %QB11 : SINT;
    ql AT %QW12 : INT;
  END_VAR
  i := k;
  arr[0] := dm;
  arr[1] := darr[0];
  arr[i] := l1;
  hs[1].r := g;
  pk(a := h.r, o => arr[2]);
  SWAP(a := arr[0], x => hs[2].r, y => tmp);
  d ?= arr[1];
  darr[1] ?= arr[0];
  qa := ID_OF(arr[0]);
  qb := ID_OF(arr[1]);
  qc := ID_OF(arr[2]);
  qd := ID_OF(hs[1].r);
  qe := ID_OF(hs[2].r);
  qf := ID_OF(tmp);
  qg := ID_OF(d);
  qh := ID_OF(darr[1]);
  qi := ID_OF(PICK(pk.o));
  tmp := darr[0].ME();
  qj := ID_OF(tmp);
  dm.GIVE(r => hs[2].r);
  qk := ID_OF(hs[2].r);
  ql := darr[0].LEVEL(pct := i * 10);
  qx0 := arr[0] = arr[1];
  qx1 := hs[1].r = rg;
  qx2 := darr[1] = NULL;
  IF stop THEN
    hs[2].r := NULL;
    hs[2].r.DAYTIME();
  END_IF;
END_PROGRAM

(* ---- itfprog.st ---- *)
(* A PROGRAM's inputs and outputs of an INTERFACE, connected in the
   CONFIGURATION (Ed.3 6.8.2) as elementary ones are: an input set from a
   global instance, from a global interface, or NULL before each run; an
   output stored into a global interface after it, a DIMMED one into a
   ROOM global. ID_OF gives a ROOM's id, 0 for NULL; gl is 2, dm 3.
   Worked by hand, k %IX0.0:
   tick 0: a gl, qa 2; b is go, NULL until the first run stores o: qb
   0; c NULL, qc 0; gr NULL until od is stored after the run, qd 0;
   o := a, so go gl; od dm, so gr dm.
   Tick 1, k TRUE: qa 2; b gl, qb 2; qd 3; o := dm, go dm.
   Tick 2, k FALSE: qb 3 (dm); o := a, go gl again.
   Tick 3: qb 2.
   reference-skip: INTERFACE and CLASS are Ed.3's, and the reference
   compiler's program connections do not compile (PROPOSAL.md §1b). *)
INTERFACE ROOM
  METHOD NAME : SINT
  END_METHOD
END_INTERFACE

INTERFACE DIMMED EXTENDS ROOM
END_INTERFACE

CLASS LIGHTROOM IMPLEMENTS ROOM
  VAR PUBLIC id : SINT; END_VAR
  METHOD PUBLIC NAME : SINT
    NAME := id;
  END_METHOD
END_CLASS

CLASS DIMMER IMPLEMENTS DIMMED
  VAR PUBLIC id : SINT; END_VAR
  METHOD PUBLIC NAME : SINT
    NAME := id;
  END_METHOD
END_CLASS

FUNCTION ID_OF : SINT
  VAR_INPUT r : ROOM; END_VAR
  IF r = NULL THEN
    ID_OF := 0;
  ELSE
    ID_OF := r.NAME();
  END_IF;
END_FUNCTION

CONFIGURATION plant
  VAR_GLOBAL
    gl : LIGHTROOM := (id := 2);
    dm : DIMMER := (id := 3);
    go : ROOM;
    gr : ROOM;
  END_VAR
  RESOURCE cpu ON PLC
    TASK fast(INTERVAL := T#10ms, PRIORITY := 1);
    PROGRAM p WITH fast : main(a := gl, b := go, c := NULL, o => go, od => gr);
  END_RESOURCE
END_CONFIGURATION

PROGRAM main
  VAR_INPUT
    a : ROOM;
    b : ROOM;
    c : ROOM;
  END_VAR
  VAR_OUTPUT
    o : ROOM;
    od : DIMMED;
  END_VAR
  VAR_EXTERNAL
    dm : DIMMER;
    gr : ROOM;
  END_VAR
  VAR
    k AT %IX0.0 : BOOL;
    qa AT %QB0 : SINT;
    qb AT %QB1 : SINT;
    qc AT %QB2 : SINT;
    qd AT %QB3 : SINT;
  END_VAR
  qa := ID_OF(a);
  qb := ID_OF(b);
  qc := ID_OF(c);
  qd := ID_OF(gr);
  IF k THEN
    o := dm;
  ELSE
    o := a;
  END_IF;
  od := dm;
END_PROGRAM

(* ---- layout2.st ---- *)
(* Structures with relative locations (Ed.3 6.4.4.7) wherever a value
   can be, and their components of other types. Worked by hand:

   Rec, 25 bytes: m, an enumeration, at 0 (starts Run, 5: 05 00); s, a
   SINT(-5..5), at 2 (starts at its lower limit -5: fb); p, a Pt, at 3
   (x 7, y -1: 07 00 ff ff); ws, a WSTRING[2] "A", at 7 (41 00, then a
   0 unit, then 0: 41 00 00 00 00 00); l, LINT -2, at 13 (fe ff ff ff ff
   ff ff ff); t, T#1s, at 21 (1000 ms: e8 03 00 00).
   V, an OVERLAP of 2 bytes: m (Mode) and w (UINT) at 0, b at bit 7 of
   byte 1; m is declared first, so it starts at Run: 05 00.

   init: gr, a global Rec at %QB0, its initial value: Q 05 00 fb 07 00
   ff ff 41 00 00 00 00 00 fe ff ff ff ff ff ff ff e8 03 00 00. img, two
   V at %QB25: 05 00 05 00. q29 0. q30 is cv.w, cv a CONSTANT V: its
   bytes, 5, not w's own initial value 0 (05).

   tick 0: the connection gives cin g's bytes (05 00) before main runs.
   a[1].p.y := 300 (2c 01), a[1].ws := "xy" (78 00 79 00 00 00), in C
   memory. fb(i := a[1], io := g): o := i, o.l := o.l * 10 = -20 (ec ff
   ff ff ff ff ff ff), io.w + 1 makes g 6 (06 00). gr := fb.o: Q0..24 05
   00 fb 07 00 2c 01 78 00 79 00 00 00 ec ff ff ff ff ff ff ff e8 03 00
   00. img[0] := cin (05 00), img[0].b := TRUE (05 80); img[1] := g (06
   00). a[0].s := 9 is clamped to 5 and flagged (CONVERSION, 4); q29 := a[0].s
   (05).

   tick 1: cin is 06 00, g 07 00 after the call: img 06 80 07 00; the
   rest as tick 0.
   reference-skip: the reference compiler (Ed.2) has no relative
   locations. *)
TYPE
  Mode : (Run := 5, Halt);
  Pt : STRUCT x : INT := 7; y : INT := -1; END_STRUCT;
  Rec : STRUCT
    m  AT %B0  : Mode;
    s  AT %B2  : SINT(-5..5);
    p  AT %B3  : Pt;
    ws AT %B7  : WSTRING[2] := "A";
    l  AT %B13 : LINT := -2;
    t  AT %B21 : TIME := T#1s;
  END_STRUCT;
  V : STRUCT OVERLAP
    m AT %B0   : Mode;
    w AT %B0   : UINT;
    b AT %X1.7 : BOOL;
  END_STRUCT;
END_TYPE
FUNCTION_BLOCK FbT
  VAR_INPUT i : Rec; END_VAR
  VAR_OUTPUT o : Rec; END_VAR
  VAR_IN_OUT io : V; END_VAR
  VAR k : Rec; END_VAR
  o := i;
  o.l := o.l * 10;
  io.w := io.w + 1;
  k.s := k.s + 1;
END_FUNCTION_BLOCK
PROGRAM main
  VAR_INPUT cin : V; END_VAR
  VAR_EXTERNAL g : V; gr : Rec; END_VAR
  VAR a : ARRAY [0..1] OF Rec; fb : FbT; END_VAR
  VAR RETAIN kept : V; END_VAR
  VAR CONSTANT cv : V; END_VAR
  VAR
    img AT %QB25 : ARRAY [0..1] OF V;
    q29 AT %QB29 : SINT;
    q30 AT %QB30 : USINT;
  END_VAR
  a[1].p.y := 300;
  a[1].ws := "xy";
  fb(i := a[1], io := g);
  gr := fb.o;
  img[0] := cin;
  img[0].b := TRUE;
  img[1] := g;
  kept := g;
  q30 := UINT_TO_USINT(cv.w);
  a[0].s := 9;
  q29 := a[0].s;
END_PROGRAM
CONFIGURATION plant
  VAR_GLOBAL
    g : V;
  END_VAR
  VAR_GLOBAL
    gr AT %QB0 : Rec;
  END_VAR
  RESOURCE r ON PLC
    TASK t (INTERVAL := T#10ms, PRIORITY := 1);
    PROGRAM p WITH t : main(cin := g);
  END_RESOURCE
END_CONFIGURATION

(* ---- locdata.st ---- *)
(* Arrays, structures and STRINGs at an address (Ed.3 6.5.5.3;
   docs/dependencies.md): from the address, their parts back to back
   with no gap, each its type's width, little-endian, a BOOL a byte, a
   STRING[n] n + 1 bytes. A structure `reading` is 11 bytes: ok at 0, raw
   at 1, at_ms at 3, label at 7. Elements read and written by computed
   index, whole arrays and structures copied in and out of the image,
   into and out of a function block, image to image, and a global at an
   address used through VAR_EXTERNAL. The initial value of `out` is
   written at the start. iecf only (reference-skip: the reference
   compiler refuses an array at an address, "Bit size of data type is
   incompatible with bit size of location", and a STRING[n] field). *)
TYPE reading :
  STRUCT
    ok : BOOL;
    raw : INT;
    at_ms : TIME;
    label : STRING[3];
  END_STRUCT;
END_TYPE

FUNCTION_BLOCK sum3
VAR_INPUT v : ARRAY[0..2] OF INT; END_VAR
VAR_OUTPUT total : INT; copy : ARRAY[0..2] OF INT; END_VAR
total := v[0] + v[1] + v[2];
copy := v;
END_FUNCTION_BLOCK

PROGRAM main
VAR
  inp AT %IW0 : ARRAY[0..2] OF INT;
  out AT %QW0 : ARRAY[0..2] OF INT := [7, 8, 9];
  flags AT %QB6 : ARRAY[0..3] OF BOOL;
  r AT %MB0 : reading;
  hist AT %MB11 : ARRAY[0..1] OF reading;
  grid AT %MB33 : ARRAY[1..2, 1..3] OF SINT;
  back AT %MW39 : ARRAY[0..2] OF INT;
END_VAR
VAR
  f : sum3;
  n, n2 : INT;
  plain : ARRAY[0..2] OF INT;
END_VAR
VAR_EXTERNAL
  gp : reading;
END_VAR
n := n + 1;
f(v := inp);
out := f.copy;
out[n MOD 3] := f.total;
r.ok := NOT r.ok;
r.raw := f.total;
r.at_ms := T#1ms * n;
IF n = 2 THEN r.label := 'xyz'; ELSE r.label := 'ab'; END_IF;
grid[2, 3] := INT_TO_SINT(n);
grid[1, n MOD 3 + 1] := -1;
hist[n MOD 2] := r;
flags[n MOD 4] := NOT flags[n MOD 4];
plain := out;
f(v := plain, total => n2, copy => back);
gp := hist[0];
END_PROGRAM

CONFIGURATION plant
  VAR_GLOBAL
    gp AT %MB45 : reading;
  END_VAR
  RESOURCE r ON PLC
    TASK fast(INTERVAL := T#10ms, PRIORITY := 0);
    PROGRAM p WITH fast : main;
  END_RESOURCE
END_CONFIGURATION
